FUNCTION "F_PressDemoCycleEnd" : Bool   // FC169, SCL
{ S7_Optimized_Access := 'TRUE' }
VERSION : 0.1
// stored: AutoNumber true, IsIECCheckEnabled false, SetENOAutomatically false, UDAEnableTagReadback false
   VAR_IN_OUT
      Seq : "FRK_SequenceCtx";
      Cycle : "ST_PressDemoCycle";
      Core : "FRK_Core";
      Unit : "FRK_Unit";
      Status : "ST_ModuleStatus";
      Part : "ST_PartContext";
      AlarmLog : "FRK_AlarmLog";
   END_VAR
   VAR_TEMP
      Written : Bool;
   END_VAR
BEGIN

   IF "FRK_SeqOnce"(Seq := #Seq, Enable := TRUE, Token := #Seq.Step) THEN
       #Cycle.CycleCompleted := TRUE;
       IF #Cycle.PartDispositioned THEN
           #Cycle.PartDispositioned := FALSE;
       ELSE
           #Written := "FRK_PartProcessed"(Core := #Core, Unit := #Unit, Status := #Status, Part := #Part, AlarmLog := #AlarmLog, Verdict := 1, Reason := 0);
           IF NOT #Written AND #Unit.CarrierIndex = 0 AND #Unit.Good < UDINT#4294967295 THEN
               #Unit.Good := #Unit.Good + 1;
           END_IF;
       END_IF;
       #Cycle.PartInMachine := FALSE;
       "FRK_SeqCycleEnd"(Seq := #Seq);
   END_IF;
   IF #Unit.StopReq THEN
       "FRK_Complete"(Core := #Core,
                      Status := #Status);
       "FRK_SeqComplete"(Seq := #Seq);
       #F_PressDemoCycleEnd := FALSE;
   ELSE
       #F_PressDemoCycleEnd := #Core.Exec <> 3;
   END_IF;
END_FUNCTION

FUNCTION_BLOCK "FB_LD_PressDemoHome"   // FB7, LAD
{ S7_Optimized_Access := 'TRUE' }
VERSION : 0.1
// stored: AutoNumber true, IsIECCheckEnabled false, IsRetainMemResEnabled false, MemoryReserve 100, SetENOAutomatically false, UDAEnableTagReadback false
   VAR_INPUT
      Run { ExternalWritable := 'False'} : Bool;
      Reset { ExternalWritable := 'False'} : Bool;
      OwnerIndex { ExternalWritable := 'False'} : DInt;
      Delta { ExternalWritable := 'False'} : Time;
   END_VAR
   VAR_IN_OUT
      PressRam : "FB_CylinderCM";
      Door : "FB_CylinderCM";
      PartSlide : "FB_CylinderCM";
   END_VAR
   VAR
      Seq { ExternalWritable := 'False'} : "FRK_SequenceCtx";
      Row1 { ExternalWritable := 'False'} : "FRK_SequenceRow";
      Row2 { ExternalWritable := 'False'} : "FRK_SequenceRow";
      Row3 { ExternalWritable := 'False'} : "FRK_SequenceRow";
      Row4 { ExternalWritable := 'False'} : "FRK_SequenceRow";
      At0 { ExternalAccessible := 'False'; ExternalVisible := 'False'; ExternalWritable := 'False'} : Bool;
      At900 { ExternalAccessible := 'False'; ExternalVisible := 'False'; ExternalWritable := 'False'} : Bool;
      At910 { ExternalAccessible := 'False'; ExternalVisible := 'False'; ExternalWritable := 'False'} : Bool;
      At999 { ExternalAccessible := 'False'; ExternalVisible := 'False'; ExternalWritable := 'False'} : Bool;
      Ready1 { ExternalAccessible := 'False'; ExternalVisible := 'False'; ExternalWritable := 'False'} : Bool;
      Ready2 { ExternalAccessible := 'False'; ExternalVisible := 'False'; ExternalWritable := 'False'} : Bool;
      Ready3 { ExternalAccessible := 'False'; ExternalVisible := 'False'; ExternalWritable := 'False'} : Bool;
      Ready4 { ExternalAccessible := 'False'; ExternalVisible := 'False'; ExternalWritable := 'False'} : Bool;
      Ready5 { ExternalAccessible := 'False'; ExternalVisible := 'False'; ExternalWritable := 'False'} : Bool;
      Advance { ExternalAccessible := 'False'; ExternalVisible := 'False'; ExternalWritable := 'False'} : Bool;
   END_VAR
BEGIN

REGION Network 1
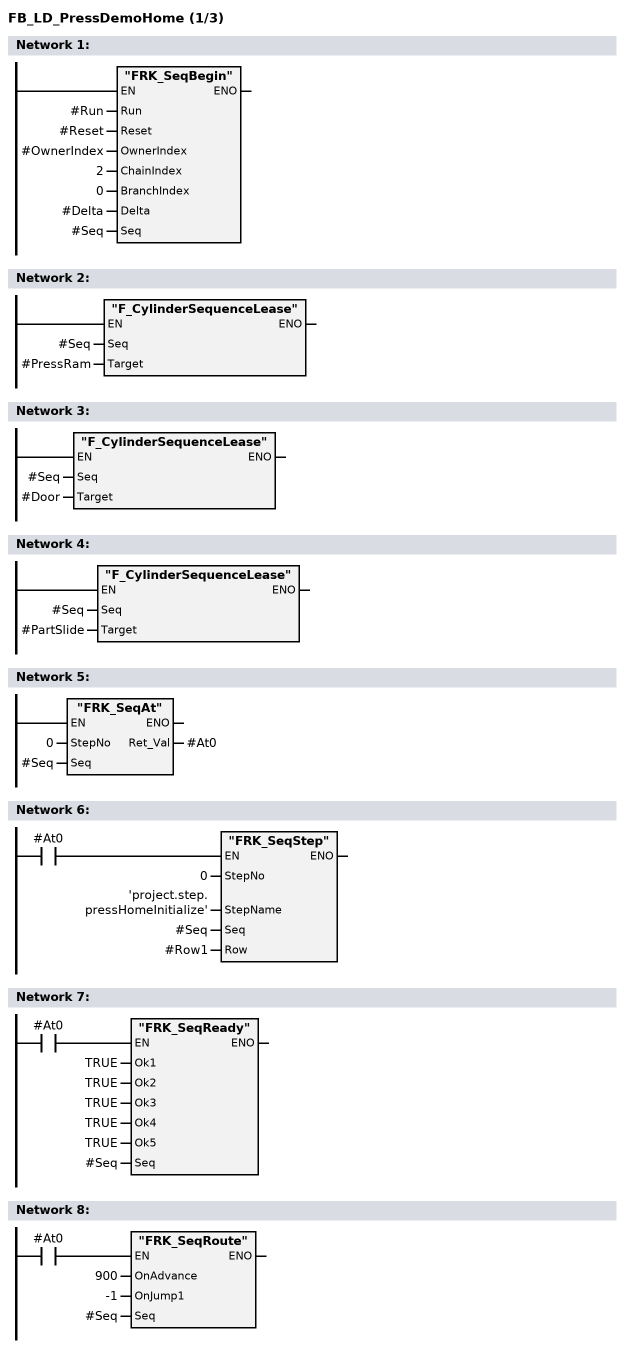
   RUNG wire#powerrail
      "FRK_SeqBegin"(Run := #Run, Reset := #Reset, OwnerIndex := #OwnerIndex, ChainIndex := 2, BranchIndex := 0, Delta := #Delta, Seq := #Seq)
   END_RUNG
   // the same network as SCL:
   "FRK_SeqBegin"(Run := #Run,
                  Reset := #Reset,
                  OwnerIndex := #OwnerIndex,
                  ChainIndex := 2,
                  BranchIndex := 0,
                  Delta := #Delta,
                  Seq := #Seq);
END_REGION

REGION Network 2
   RUNG wire#powerrail
      "F_CylinderSequenceLease"(Seq := #Seq, Target := #PressRam)
   END_RUNG
   // the same network as SCL:
   "F_CylinderSequenceLease"(Seq := #Seq, Target := #PressRam);
END_REGION

REGION Network 3
   RUNG wire#powerrail
      "F_CylinderSequenceLease"(Seq := #Seq, Target := #Door)
   END_RUNG
   // the same network as SCL:
   "F_CylinderSequenceLease"(Seq := #Seq, Target := #Door);
END_REGION

REGION Network 4
   RUNG wire#powerrail
      "F_CylinderSequenceLease"(Seq := #Seq, Target := #PartSlide)
   END_RUNG
   // the same network as SCL:
   "F_CylinderSequenceLease"(Seq := #Seq, Target := #PartSlide);
END_REGION

REGION Network 5
   RUNG wire#powerrail
      "FRK_SeqAt"(StepNo := 0, Seq := #Seq, Ret_Val => #At0)
   END_RUNG
   // the same network as SCL:
   #At0 := "FRK_SeqAt"(StepNo := 0, Seq := #Seq);
END_REGION

REGION Network 6
   RUNG wire#powerrail
      Contact( #At0 )
      "FRK_SeqStep"(StepNo := 0, StepName := 'project.step.pressHomeInitialize', Seq := #Seq, Row := #Row1)
   END_RUNG
   // the same network as SCL:
   IF #At0 THEN
       "FRK_SeqStep"(StepNo := 0, StepName := 'project.step.pressHomeInitialize', Seq := #Seq, Row := #Row1);
   END_IF;
END_REGION

REGION Network 7
   RUNG wire#powerrail
      Contact( #At0 )
      "FRK_SeqReady"(Ok1 := TRUE, Ok2 := TRUE, Ok3 := TRUE, Ok4 := TRUE, Ok5 := TRUE, Seq := #Seq)
   END_RUNG
   // the same network as SCL:
   IF #At0 THEN
       "FRK_SeqReady"(Ok1 := TRUE, Ok2 := TRUE, Ok3 := TRUE, Ok4 := TRUE, Ok5 := TRUE, Seq := #Seq);
   END_IF;
END_REGION

REGION Network 8
   RUNG wire#powerrail
      Contact( #At0 )
      "FRK_SeqRoute"(OnAdvance := 900, OnJump1 := -1, Seq := #Seq)
   END_RUNG
   // the same network as SCL:
   IF #At0 THEN "FRK_SeqRoute"(OnAdvance := 900, OnJump1 := -1, Seq := #Seq); END_IF;
END_REGION

REGION Network 9
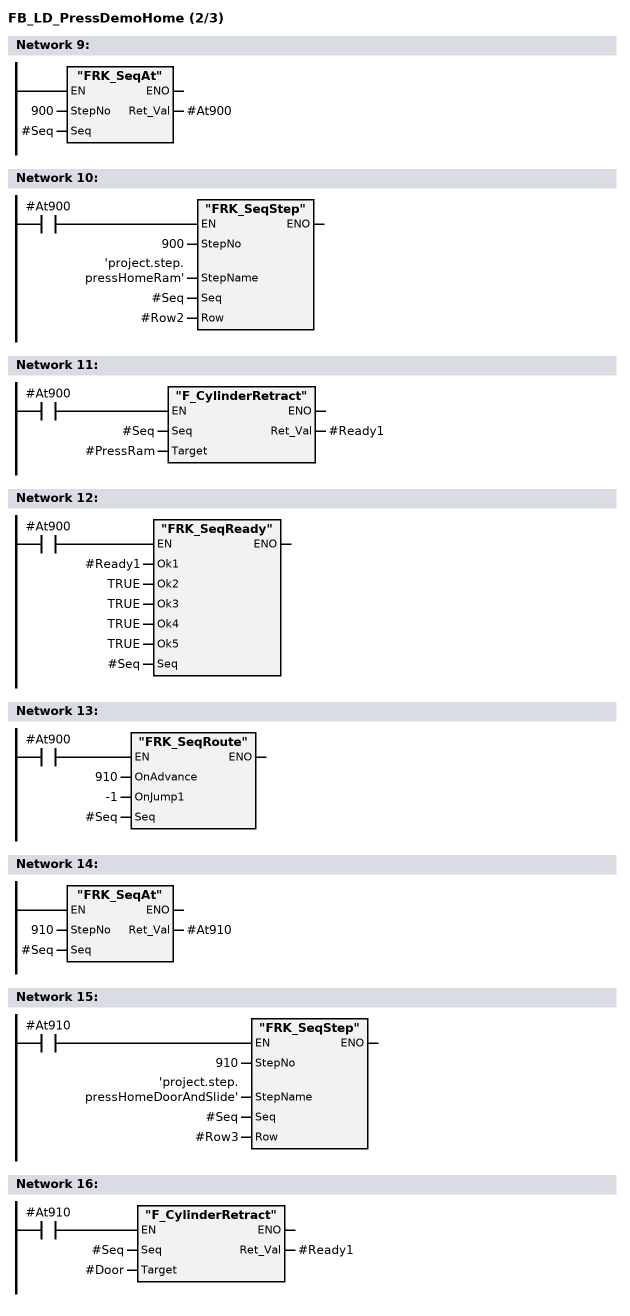
   RUNG wire#powerrail
      "FRK_SeqAt"(StepNo := 900, Seq := #Seq, Ret_Val => #At900)
   END_RUNG
   // the same network as SCL:
   #At900 := "FRK_SeqAt"(StepNo := 900, Seq := #Seq);
END_REGION

REGION Network 10
   RUNG wire#powerrail
      Contact( #At900 )
      "FRK_SeqStep"(StepNo := 900, StepName := 'project.step.pressHomeRam', Seq := #Seq, Row := #Row2)
   END_RUNG
   // the same network as SCL:
   IF #At900 THEN
       "FRK_SeqStep"(StepNo := 900, StepName := 'project.step.pressHomeRam', Seq := #Seq, Row := #Row2);
   END_IF;
END_REGION

REGION Network 11
   RUNG wire#powerrail
      Contact( #At900 )
      "F_CylinderRetract"(Seq := #Seq, Target := #PressRam, Ret_Val => #Ready1)
   END_RUNG
   // the same network as SCL:
   IF #At900 THEN #Ready1 := "F_CylinderRetract"(Seq := #Seq, Target := #PressRam); END_IF;
END_REGION

REGION Network 12
   RUNG wire#powerrail
      Contact( #At900 )
      "FRK_SeqReady"(Ok1 := #Ready1, Ok2 := TRUE, Ok3 := TRUE, Ok4 := TRUE, Ok5 := TRUE, Seq := #Seq)
   END_RUNG
   // the same network as SCL:
   IF #At900 THEN
       "FRK_SeqReady"(Ok1 := #Ready1, Ok2 := TRUE, Ok3 := TRUE, Ok4 := TRUE, Ok5 := TRUE, Seq := #Seq);
   END_IF;
END_REGION

REGION Network 13
   RUNG wire#powerrail
      Contact( #At900 )
      "FRK_SeqRoute"(OnAdvance := 910, OnJump1 := -1, Seq := #Seq)
   END_RUNG
   // the same network as SCL:
   IF #At900 THEN "FRK_SeqRoute"(OnAdvance := 910, OnJump1 := -1, Seq := #Seq); END_IF;
END_REGION

REGION Network 14
   RUNG wire#powerrail
      "FRK_SeqAt"(StepNo := 910, Seq := #Seq, Ret_Val => #At910)
   END_RUNG
   // the same network as SCL:
   #At910 := "FRK_SeqAt"(StepNo := 910, Seq := #Seq);
END_REGION

REGION Network 15
   RUNG wire#powerrail
      Contact( #At910 )
      "FRK_SeqStep"(StepNo := 910, StepName := 'project.step.pressHomeDoorAndSlide', Seq := #Seq, Row := #Row3)
   END_RUNG
   // the same network as SCL:
   IF #At910 THEN
       "FRK_SeqStep"(StepNo := 910, StepName := 'project.step.pressHomeDoorAndSlide', Seq := #Seq, Row := #Row3);
   END_IF;
END_REGION

REGION Network 16
   RUNG wire#powerrail
      Contact( #At910 )
      "F_CylinderRetract"(Seq := #Seq, Target := #Door, Ret_Val => #Ready1)
   END_RUNG
   // the same network as SCL:
   IF #At910 THEN #Ready1 := "F_CylinderRetract"(Seq := #Seq, Target := #Door); END_IF;
END_REGION

REGION Network 17
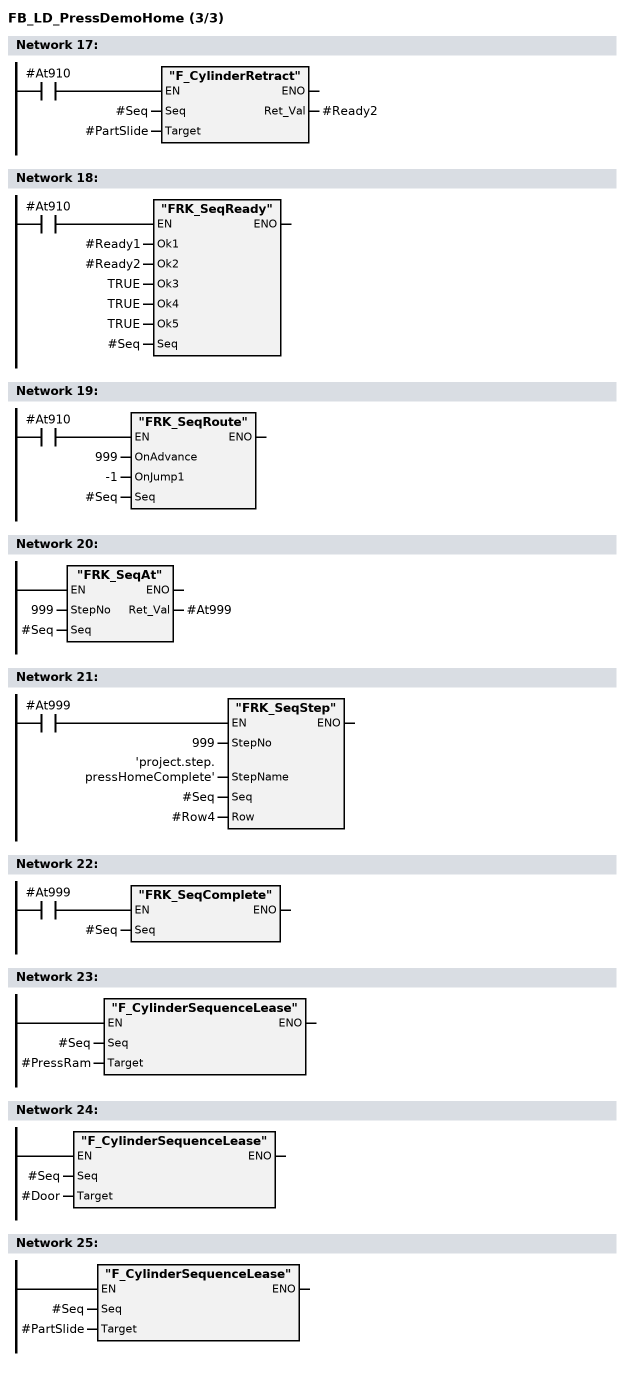
   RUNG wire#powerrail
      Contact( #At910 )
      "F_CylinderRetract"(Seq := #Seq, Target := #PartSlide, Ret_Val => #Ready2)
   END_RUNG
   // the same network as SCL:
   IF #At910 THEN #Ready2 := "F_CylinderRetract"(Seq := #Seq, Target := #PartSlide); END_IF;
END_REGION

REGION Network 18
   RUNG wire#powerrail
      Contact( #At910 )
      "FRK_SeqReady"(Ok1 := #Ready1, Ok2 := #Ready2, Ok3 := TRUE, Ok4 := TRUE, Ok5 := TRUE, Seq := #Seq)
   END_RUNG
   // the same network as SCL:
   IF #At910 THEN
       "FRK_SeqReady"(Ok1 := #Ready1, Ok2 := #Ready2, Ok3 := TRUE, Ok4 := TRUE, Ok5 := TRUE, Seq := #Seq);
   END_IF;
END_REGION

REGION Network 19
   RUNG wire#powerrail
      Contact( #At910 )
      "FRK_SeqRoute"(OnAdvance := 999, OnJump1 := -1, Seq := #Seq)
   END_RUNG
   // the same network as SCL:
   IF #At910 THEN "FRK_SeqRoute"(OnAdvance := 999, OnJump1 := -1, Seq := #Seq); END_IF;
END_REGION

REGION Network 20
   RUNG wire#powerrail
      "FRK_SeqAt"(StepNo := 999, Seq := #Seq, Ret_Val => #At999)
   END_RUNG
   // the same network as SCL:
   #At999 := "FRK_SeqAt"(StepNo := 999, Seq := #Seq);
END_REGION

REGION Network 21
   RUNG wire#powerrail
      Contact( #At999 )
      "FRK_SeqStep"(StepNo := 999, StepName := 'project.step.pressHomeComplete', Seq := #Seq, Row := #Row4)
   END_RUNG
   // the same network as SCL:
   IF #At999 THEN
       "FRK_SeqStep"(StepNo := 999, StepName := 'project.step.pressHomeComplete', Seq := #Seq, Row := #Row4);
   END_IF;
END_REGION

REGION Network 22
   RUNG wire#powerrail
      Contact( #At999 )
      "FRK_SeqComplete"(Seq := #Seq)
   END_RUNG
   // the same network as SCL:
   IF #At999 THEN "FRK_SeqComplete"(Seq := #Seq); END_IF;
END_REGION

REGION Network 23
   RUNG wire#powerrail
      "F_CylinderSequenceLease"(Seq := #Seq, Target := #PressRam)
   END_RUNG
   // the same network as SCL:
   "F_CylinderSequenceLease"(Seq := #Seq, Target := #PressRam);
END_REGION

REGION Network 24
   RUNG wire#powerrail
      "F_CylinderSequenceLease"(Seq := #Seq, Target := #Door)
   END_RUNG
   // the same network as SCL:
   "F_CylinderSequenceLease"(Seq := #Seq, Target := #Door);
END_REGION

REGION Network 25
   RUNG wire#powerrail
      "F_CylinderSequenceLease"(Seq := #Seq, Target := #PartSlide)
   END_RUNG
   // the same network as SCL:
   "F_CylinderSequenceLease"(Seq := #Seq, Target := #PartSlide);
END_REGION
END_FUNCTION_BLOCK

FUNCTION "FRK_SeqComplete" : Void   // FC127, SCL
{ S7_Optimized_Access := 'TRUE' }
VERSION : 0.1
// stored: AutoNumber true, IsIECCheckEnabled false, SetENOAutomatically false, UDAEnableTagReadback false
   VAR_IN_OUT
      Seq : "FRK_SequenceCtx";
   END_VAR
BEGIN

   #Seq.Done := TRUE;
   #Seq.Running := FALSE;
END_FUNCTION

FUNCTION_BLOCK "FB_LD_PressDemoLoadPosition"   // FB8, LAD
{ S7_Optimized_Access := 'TRUE' }
VERSION : 0.1
// stored: AutoNumber true, IsIECCheckEnabled false, IsRetainMemResEnabled false, MemoryReserve 100, SetENOAutomatically false, UDAEnableTagReadback false
   VAR_INPUT
      Run { ExternalWritable := 'False'} : Bool;
      Reset { ExternalWritable := 'False'} : Bool;
      OwnerIndex { ExternalWritable := 'False'} : DInt;
      Delta { ExternalWritable := 'False'} : Time;
   END_VAR
   VAR_IN_OUT
      PressRam : "FB_CylinderCM";
      Door : "FB_CylinderCM";
      PartSlide : "FB_CylinderCM";
   END_VAR
   VAR
      Seq { ExternalWritable := 'False'} : "FRK_SequenceCtx";
      Row1 { ExternalWritable := 'False'} : "FRK_SequenceRow";
      Row2 { ExternalWritable := 'False'} : "FRK_SequenceRow";
      Row3 { ExternalWritable := 'False'} : "FRK_SequenceRow";
      Row4 { ExternalWritable := 'False'} : "FRK_SequenceRow";
      At240 { ExternalAccessible := 'False'; ExternalVisible := 'False'; ExternalWritable := 'False'} : Bool;
      At260 { ExternalAccessible := 'False'; ExternalVisible := 'False'; ExternalWritable := 'False'} : Bool;
      At280 { ExternalAccessible := 'False'; ExternalVisible := 'False'; ExternalWritable := 'False'} : Bool;
      At300 { ExternalAccessible := 'False'; ExternalVisible := 'False'; ExternalWritable := 'False'} : Bool;
      Ready1 { ExternalAccessible := 'False'; ExternalVisible := 'False'; ExternalWritable := 'False'} : Bool;
      Ready2 { ExternalAccessible := 'False'; ExternalVisible := 'False'; ExternalWritable := 'False'} : Bool;
      Ready3 { ExternalAccessible := 'False'; ExternalVisible := 'False'; ExternalWritable := 'False'} : Bool;
      Ready4 { ExternalAccessible := 'False'; ExternalVisible := 'False'; ExternalWritable := 'False'} : Bool;
      Ready5 { ExternalAccessible := 'False'; ExternalVisible := 'False'; ExternalWritable := 'False'} : Bool;
      Advance { ExternalAccessible := 'False'; ExternalVisible := 'False'; ExternalWritable := 'False'} : Bool;
   END_VAR
BEGIN

REGION Network 1
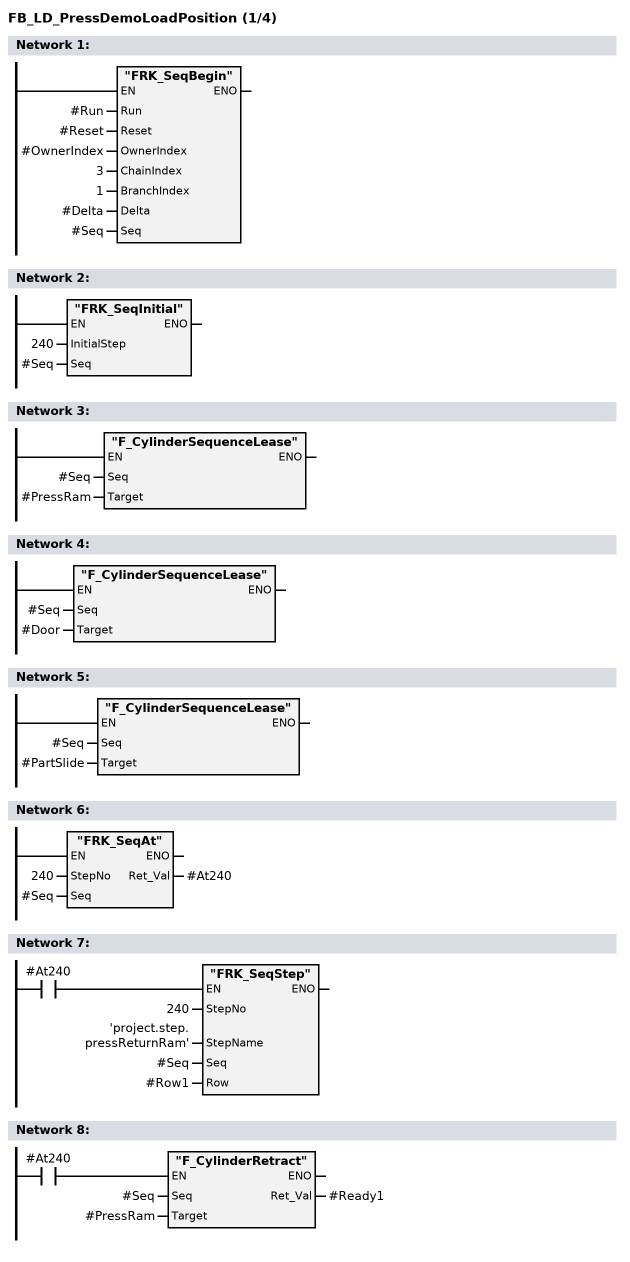
   RUNG wire#powerrail
      "FRK_SeqBegin"(Run := #Run, Reset := #Reset, OwnerIndex := #OwnerIndex, ChainIndex := 3, BranchIndex := 1, Delta := #Delta, Seq := #Seq)
   END_RUNG
   // the same network as SCL:
   "FRK_SeqBegin"(Run := #Run,
                  Reset := #Reset,
                  OwnerIndex := #OwnerIndex,
                  ChainIndex := 3,
                  BranchIndex := 1,
                  Delta := #Delta,
                  Seq := #Seq);
END_REGION

REGION Network 2
   RUNG wire#powerrail
      "FRK_SeqInitial"(InitialStep := 240, Seq := #Seq)
   END_RUNG
   // the same network as SCL:
   "FRK_SeqInitial"(InitialStep := 240, Seq := #Seq);
END_REGION

REGION Network 3
   RUNG wire#powerrail
      "F_CylinderSequenceLease"(Seq := #Seq, Target := #PressRam)
   END_RUNG
   // the same network as SCL:
   "F_CylinderSequenceLease"(Seq := #Seq, Target := #PressRam);
END_REGION

REGION Network 4
   RUNG wire#powerrail
      "F_CylinderSequenceLease"(Seq := #Seq, Target := #Door)
   END_RUNG
   // the same network as SCL:
   "F_CylinderSequenceLease"(Seq := #Seq, Target := #Door);
END_REGION

REGION Network 5
   RUNG wire#powerrail
      "F_CylinderSequenceLease"(Seq := #Seq, Target := #PartSlide)
   END_RUNG
   // the same network as SCL:
   "F_CylinderSequenceLease"(Seq := #Seq, Target := #PartSlide);
END_REGION

REGION Network 6
   RUNG wire#powerrail
      "FRK_SeqAt"(StepNo := 240, Seq := #Seq, Ret_Val => #At240)
   END_RUNG
   // the same network as SCL:
   #At240 := "FRK_SeqAt"(StepNo := 240, Seq := #Seq);
END_REGION

REGION Network 7
   RUNG wire#powerrail
      Contact( #At240 )
      "FRK_SeqStep"(StepNo := 240, StepName := 'project.step.pressReturnRam', Seq := #Seq, Row := #Row1)
   END_RUNG
   // the same network as SCL:
   IF #At240 THEN
       "FRK_SeqStep"(StepNo := 240, StepName := 'project.step.pressReturnRam', Seq := #Seq, Row := #Row1);
   END_IF;
END_REGION

REGION Network 8
   RUNG wire#powerrail
      Contact( #At240 )
      "F_CylinderRetract"(Seq := #Seq, Target := #PressRam, Ret_Val => #Ready1)
   END_RUNG
   // the same network as SCL:
   IF #At240 THEN #Ready1 := "F_CylinderRetract"(Seq := #Seq, Target := #PressRam); END_IF;
END_REGION

REGION Network 9
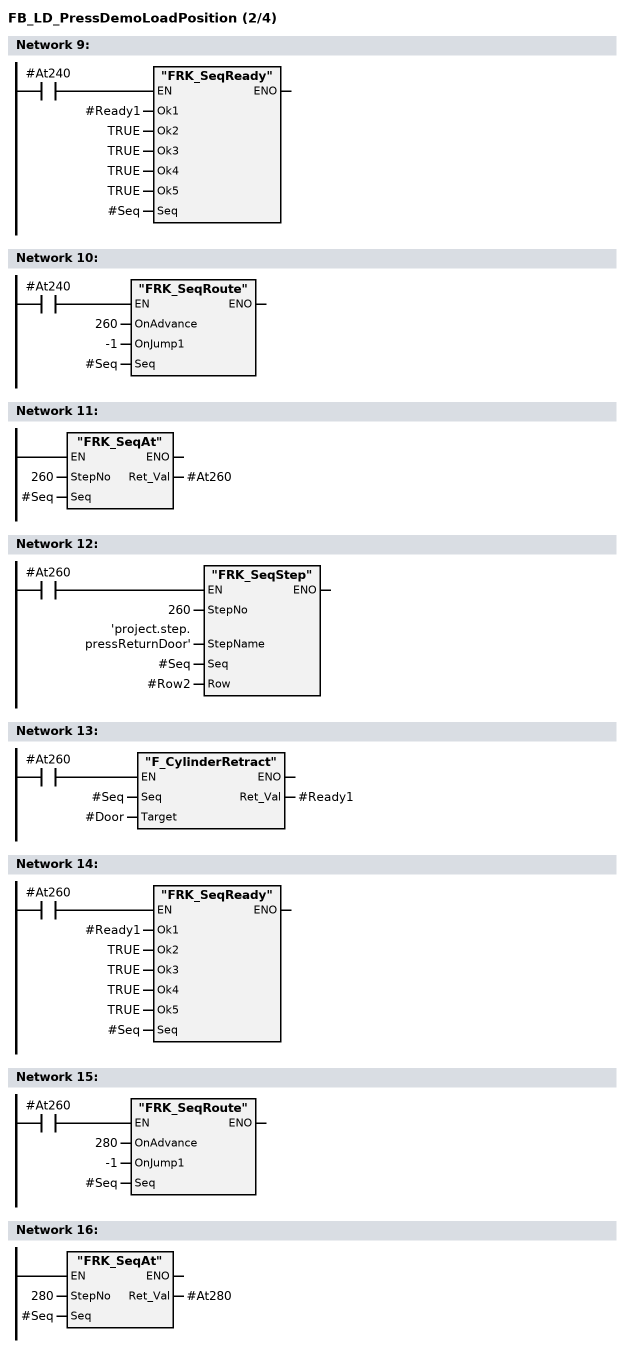
   RUNG wire#powerrail
      Contact( #At240 )
      "FRK_SeqReady"(Ok1 := #Ready1, Ok2 := TRUE, Ok3 := TRUE, Ok4 := TRUE, Ok5 := TRUE, Seq := #Seq)
   END_RUNG
   // the same network as SCL:
   IF #At240 THEN
       "FRK_SeqReady"(Ok1 := #Ready1, Ok2 := TRUE, Ok3 := TRUE, Ok4 := TRUE, Ok5 := TRUE, Seq := #Seq);
   END_IF;
END_REGION

REGION Network 10
   RUNG wire#powerrail
      Contact( #At240 )
      "FRK_SeqRoute"(OnAdvance := 260, OnJump1 := -1, Seq := #Seq)
   END_RUNG
   // the same network as SCL:
   IF #At240 THEN "FRK_SeqRoute"(OnAdvance := 260, OnJump1 := -1, Seq := #Seq); END_IF;
END_REGION

REGION Network 11
   RUNG wire#powerrail
      "FRK_SeqAt"(StepNo := 260, Seq := #Seq, Ret_Val => #At260)
   END_RUNG
   // the same network as SCL:
   #At260 := "FRK_SeqAt"(StepNo := 260, Seq := #Seq);
END_REGION

REGION Network 12
   RUNG wire#powerrail
      Contact( #At260 )
      "FRK_SeqStep"(StepNo := 260, StepName := 'project.step.pressReturnDoor', Seq := #Seq, Row := #Row2)
   END_RUNG
   // the same network as SCL:
   IF #At260 THEN
       "FRK_SeqStep"(StepNo := 260, StepName := 'project.step.pressReturnDoor', Seq := #Seq, Row := #Row2);
   END_IF;
END_REGION

REGION Network 13
   RUNG wire#powerrail
      Contact( #At260 )
      "F_CylinderRetract"(Seq := #Seq, Target := #Door, Ret_Val => #Ready1)
   END_RUNG
   // the same network as SCL:
   IF #At260 THEN #Ready1 := "F_CylinderRetract"(Seq := #Seq, Target := #Door); END_IF;
END_REGION

REGION Network 14
   RUNG wire#powerrail
      Contact( #At260 )
      "FRK_SeqReady"(Ok1 := #Ready1, Ok2 := TRUE, Ok3 := TRUE, Ok4 := TRUE, Ok5 := TRUE, Seq := #Seq)
   END_RUNG
   // the same network as SCL:
   IF #At260 THEN
       "FRK_SeqReady"(Ok1 := #Ready1, Ok2 := TRUE, Ok3 := TRUE, Ok4 := TRUE, Ok5 := TRUE, Seq := #Seq);
   END_IF;
END_REGION

REGION Network 15
   RUNG wire#powerrail
      Contact( #At260 )
      "FRK_SeqRoute"(OnAdvance := 280, OnJump1 := -1, Seq := #Seq)
   END_RUNG
   // the same network as SCL:
   IF #At260 THEN "FRK_SeqRoute"(OnAdvance := 280, OnJump1 := -1, Seq := #Seq); END_IF;
END_REGION

REGION Network 16
   RUNG wire#powerrail
      "FRK_SeqAt"(StepNo := 280, Seq := #Seq, Ret_Val => #At280)
   END_RUNG
   // the same network as SCL:
   #At280 := "FRK_SeqAt"(StepNo := 280, Seq := #Seq);
END_REGION

REGION Network 17
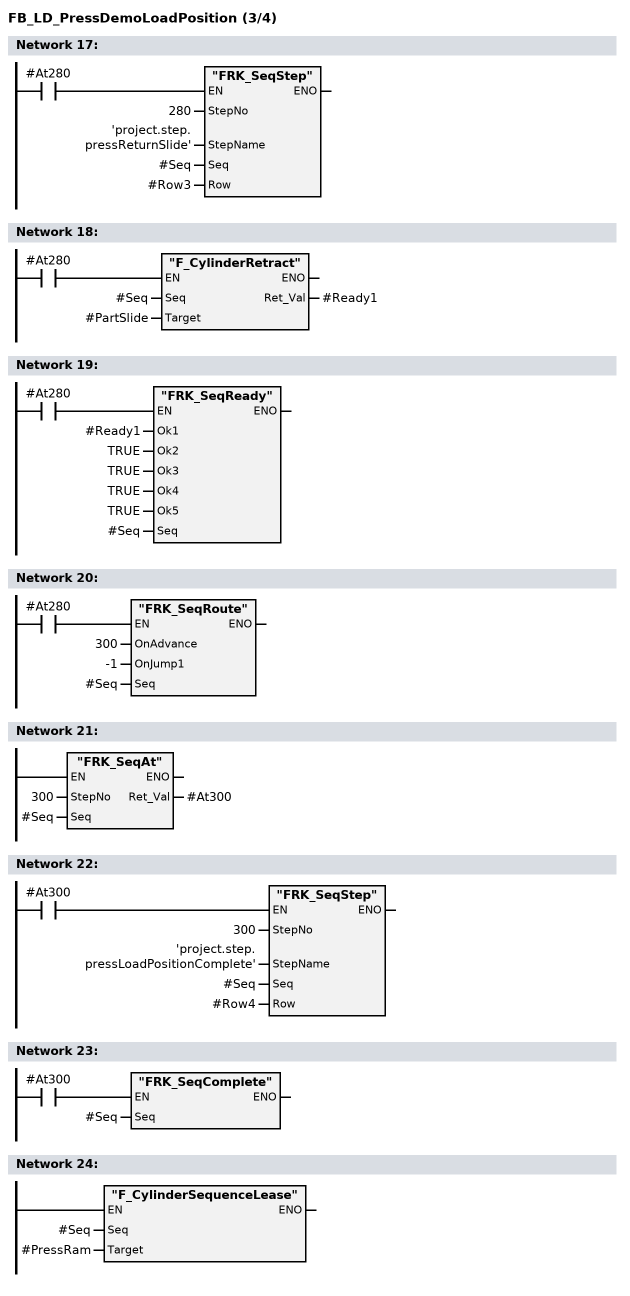
   RUNG wire#powerrail
      Contact( #At280 )
      "FRK_SeqStep"(StepNo := 280, StepName := 'project.step.pressReturnSlide', Seq := #Seq, Row := #Row3)
   END_RUNG
   // the same network as SCL:
   IF #At280 THEN
       "FRK_SeqStep"(StepNo := 280, StepName := 'project.step.pressReturnSlide', Seq := #Seq, Row := #Row3);
   END_IF;
END_REGION

REGION Network 18
   RUNG wire#powerrail
      Contact( #At280 )
      "F_CylinderRetract"(Seq := #Seq, Target := #PartSlide, Ret_Val => #Ready1)
   END_RUNG
   // the same network as SCL:
   IF #At280 THEN #Ready1 := "F_CylinderRetract"(Seq := #Seq, Target := #PartSlide); END_IF;
END_REGION

REGION Network 19
   RUNG wire#powerrail
      Contact( #At280 )
      "FRK_SeqReady"(Ok1 := #Ready1, Ok2 := TRUE, Ok3 := TRUE, Ok4 := TRUE, Ok5 := TRUE, Seq := #Seq)
   END_RUNG
   // the same network as SCL:
   IF #At280 THEN
       "FRK_SeqReady"(Ok1 := #Ready1, Ok2 := TRUE, Ok3 := TRUE, Ok4 := TRUE, Ok5 := TRUE, Seq := #Seq);
   END_IF;
END_REGION

REGION Network 20
   RUNG wire#powerrail
      Contact( #At280 )
      "FRK_SeqRoute"(OnAdvance := 300, OnJump1 := -1, Seq := #Seq)
   END_RUNG
   // the same network as SCL:
   IF #At280 THEN "FRK_SeqRoute"(OnAdvance := 300, OnJump1 := -1, Seq := #Seq); END_IF;
END_REGION

REGION Network 21
   RUNG wire#powerrail
      "FRK_SeqAt"(StepNo := 300, Seq := #Seq, Ret_Val => #At300)
   END_RUNG
   // the same network as SCL:
   #At300 := "FRK_SeqAt"(StepNo := 300, Seq := #Seq);
END_REGION

REGION Network 22
   RUNG wire#powerrail
      Contact( #At300 )
      "FRK_SeqStep"(StepNo := 300, StepName := 'project.step.pressLoadPositionComplete', Seq := #Seq, Row := #Row4)
   END_RUNG
   // the same network as SCL:
   IF #At300 THEN
       "FRK_SeqStep"(StepNo := 300, StepName := 'project.step.pressLoadPositionComplete', Seq := #Seq, Row := #Row4);
   END_IF;
END_REGION

REGION Network 23
   RUNG wire#powerrail
      Contact( #At300 )
      "FRK_SeqComplete"(Seq := #Seq)
   END_RUNG
   // the same network as SCL:
   IF #At300 THEN "FRK_SeqComplete"(Seq := #Seq); END_IF;
END_REGION

REGION Network 24
   RUNG wire#powerrail
      "F_CylinderSequenceLease"(Seq := #Seq, Target := #PressRam)
   END_RUNG
   // the same network as SCL:
   "F_CylinderSequenceLease"(Seq := #Seq, Target := #PressRam);
END_REGION

REGION Network 25
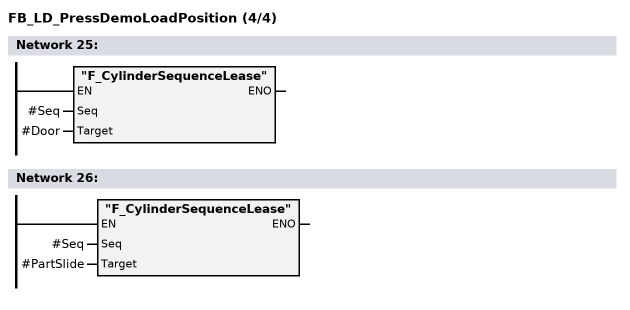
   RUNG wire#powerrail
      "F_CylinderSequenceLease"(Seq := #Seq, Target := #Door)
   END_RUNG
   // the same network as SCL:
   "F_CylinderSequenceLease"(Seq := #Seq, Target := #Door);
END_REGION

REGION Network 26
   RUNG wire#powerrail
      "F_CylinderSequenceLease"(Seq := #Seq, Target := #PartSlide)
   END_RUNG
   // the same network as SCL:
   "F_CylinderSequenceLease"(Seq := #Seq, Target := #PartSlide);
END_REGION
END_FUNCTION_BLOCK

FUNCTION "FRK_SeqInitial" : Void   // FC135, SCL
{ S7_Optimized_Access := 'TRUE' }
VERSION : 0.1
// stored: AutoNumber true, IsIECCheckEnabled false, SetENOAutomatically false, UDAEnableTagReadback false
   VAR_INPUT
      InitialStep : DInt;
   END_VAR
   VAR_IN_OUT
      Seq : "FRK_SequenceCtx";
   END_VAR
BEGIN

   IF #Seq.Restart OR NOT #Seq.Running THEN
       #Seq.Step := #InitialStep;
       #Seq.ScanStep := #InitialStep;
   END_IF;
END_FUNCTION

FUNCTION_BLOCK "FB_LD_PressDemoRelease"   // FB9, LAD
{ S7_Optimized_Access := 'TRUE' }
VERSION : 0.1
// stored: AutoNumber true, IsIECCheckEnabled false, IsRetainMemResEnabled false, MemoryReserve 100, SetENOAutomatically false, UDAEnableTagReadback false
   VAR_INPUT
      AirPressureOk { ExternalWritable := 'False'} : Bool;
      DoorClosed { ExternalWritable := 'False'} : Bool;
      DoorHealthy { ExternalWritable := 'False'} : Bool;
      RamHealthy { ExternalWritable := 'False'} : Bool;
      SlideHealthy { ExternalWritable := 'False'} : Bool;
      SlideInside { ExternalWritable := 'False'} : Bool;
      TwoHandHeld { ExternalWritable := 'False'} : Bool;
   END_VAR
   VAR
      Conditions { ExternalWritable := 'False'} : "ST_PressDemoReleaseConditions";
      ModeStart { ExternalWritable := 'False'} : "FRK_PermCtx";
      RamExtend { ExternalWritable := 'False'} : "FRK_PermCtx";
   END_VAR
BEGIN

REGION Network 1
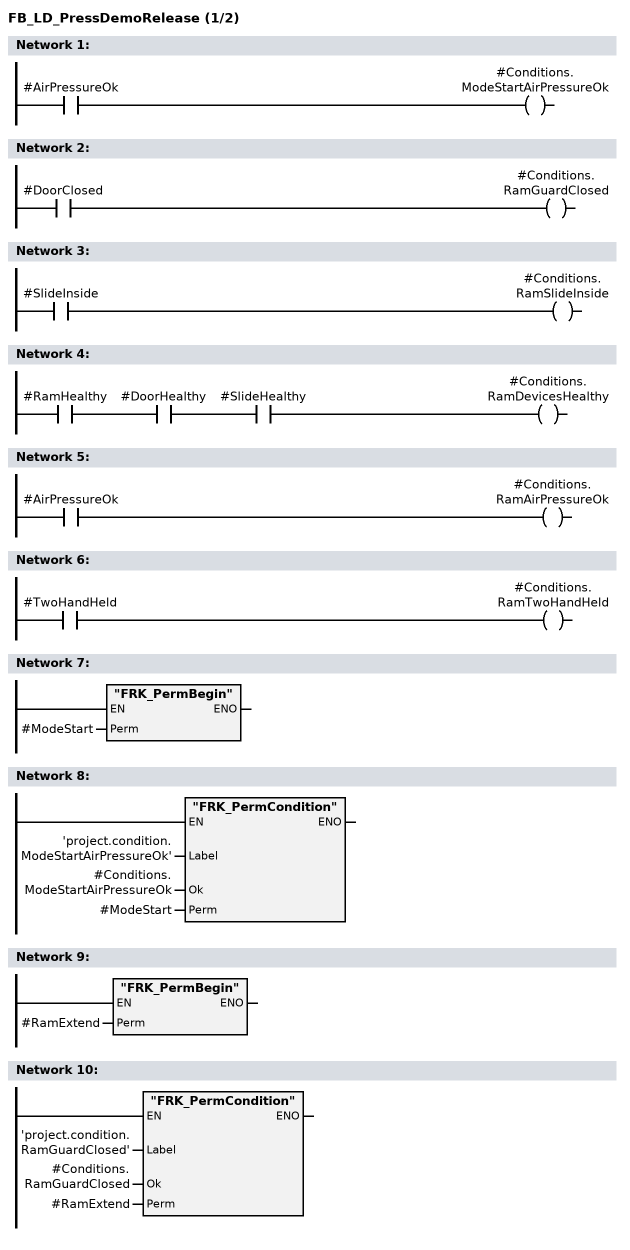
   RUNG wire#powerrail
      Contact( #AirPressureOk )
      Coil( #Conditions.ModeStartAirPressureOk )
   END_RUNG
   // the same network as SCL:
   #Conditions.ModeStartAirPressureOk := #AirPressureOk;
END_REGION

REGION Network 2
   RUNG wire#powerrail
      Contact( #DoorClosed )
      Coil( #Conditions.RamGuardClosed )
   END_RUNG
   // the same network as SCL:
   #Conditions.RamGuardClosed := #DoorClosed;
END_REGION

REGION Network 3
   RUNG wire#powerrail
      Contact( #SlideInside )
      Coil( #Conditions.RamSlideInside )
   END_RUNG
   // the same network as SCL:
   #Conditions.RamSlideInside := #SlideInside;
END_REGION

REGION Network 4
   RUNG wire#powerrail
      Contact( #RamHealthy )
      Contact( #DoorHealthy )
      Contact( #SlideHealthy )
      Coil( #Conditions.RamDevicesHealthy )
   END_RUNG
   // the same network as SCL:
   #Conditions.RamDevicesHealthy := #RamHealthy AND #DoorHealthy AND #SlideHealthy;
END_REGION

REGION Network 5
   RUNG wire#powerrail
      Contact( #AirPressureOk )
      Coil( #Conditions.RamAirPressureOk )
   END_RUNG
   // the same network as SCL:
   #Conditions.RamAirPressureOk := #AirPressureOk;
END_REGION

REGION Network 6
   RUNG wire#powerrail
      Contact( #TwoHandHeld )
      Coil( #Conditions.RamTwoHandHeld )
   END_RUNG
   // the same network as SCL:
   #Conditions.RamTwoHandHeld := #TwoHandHeld;
END_REGION

REGION Network 7
   RUNG wire#powerrail
      "FRK_PermBegin"(Perm := #ModeStart)
   END_RUNG
   // the same network as SCL:
   "FRK_PermBegin"(Perm := #ModeStart);
END_REGION

REGION Network 8
   RUNG wire#powerrail
      "FRK_PermCondition"(Label := 'project.condition.ModeStartAirPressureOk', Ok := #Conditions.ModeStartAirPressureOk, Perm := #ModeStart)
   END_RUNG
   // the same network as SCL:
   "FRK_PermCondition"(Label := 'project.condition.ModeStartAirPressureOk',
                       Ok := #Conditions.ModeStartAirPressureOk,
                       Perm := #ModeStart);
END_REGION

REGION Network 9
   RUNG wire#powerrail
      "FRK_PermBegin"(Perm := #RamExtend)
   END_RUNG
   // the same network as SCL:
   "FRK_PermBegin"(Perm := #RamExtend);
END_REGION

REGION Network 10
   RUNG wire#powerrail
      "FRK_PermCondition"(Label := 'project.condition.RamGuardClosed', Ok := #Conditions.RamGuardClosed, Perm := #RamExtend)
   END_RUNG
   // the same network as SCL:
   "FRK_PermCondition"(Label := 'project.condition.RamGuardClosed',
                       Ok := #Conditions.RamGuardClosed,
                       Perm := #RamExtend);
END_REGION

REGION Network 11
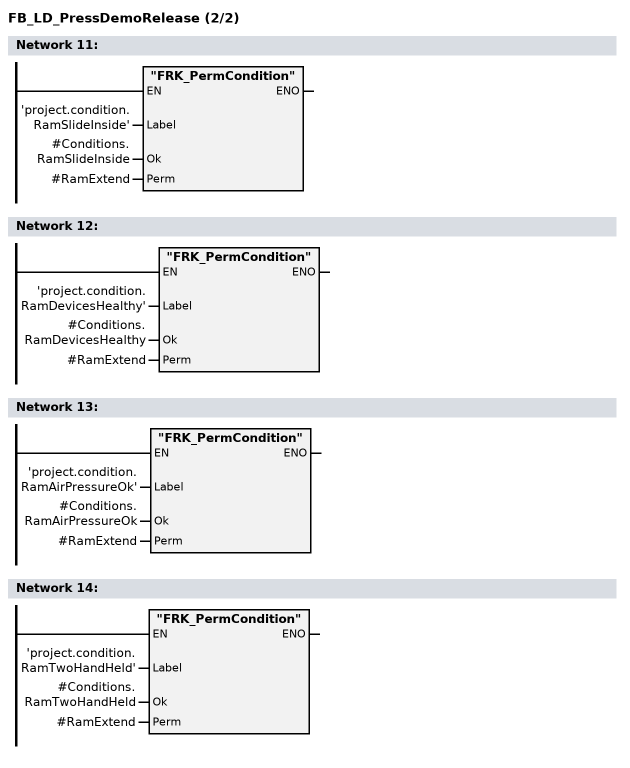
   RUNG wire#powerrail
      "FRK_PermCondition"(Label := 'project.condition.RamSlideInside', Ok := #Conditions.RamSlideInside, Perm := #RamExtend)
   END_RUNG
   // the same network as SCL:
   "FRK_PermCondition"(Label := 'project.condition.RamSlideInside',
                       Ok := #Conditions.RamSlideInside,
                       Perm := #RamExtend);
END_REGION

REGION Network 12
   RUNG wire#powerrail
      "FRK_PermCondition"(Label := 'project.condition.RamDevicesHealthy', Ok := #Conditions.RamDevicesHealthy, Perm := #RamExtend)
   END_RUNG
   // the same network as SCL:
   "FRK_PermCondition"(Label := 'project.condition.RamDevicesHealthy',
                       Ok := #Conditions.RamDevicesHealthy,
                       Perm := #RamExtend);
END_REGION

REGION Network 13
   RUNG wire#powerrail
      "FRK_PermCondition"(Label := 'project.condition.RamAirPressureOk', Ok := #Conditions.RamAirPressureOk, Perm := #RamExtend)
   END_RUNG
   // the same network as SCL:
   "FRK_PermCondition"(Label := 'project.condition.RamAirPressureOk',
                       Ok := #Conditions.RamAirPressureOk,
                       Perm := #RamExtend);
END_REGION

REGION Network 14
   RUNG wire#powerrail
      "FRK_PermCondition"(Label := 'project.condition.RamTwoHandHeld', Ok := #Conditions.RamTwoHandHeld, Perm := #RamExtend)
   END_RUNG
   // the same network as SCL:
   "FRK_PermCondition"(Label := 'project.condition.RamTwoHandHeld',
                       Ok := #Conditions.RamTwoHandHeld,
                       Perm := #RamExtend);
END_REGION
END_FUNCTION_BLOCK

FUNCTION "FRK_PermBegin" : Void   // FC122, SCL
{ S7_Optimized_Access := 'TRUE' }
VERSION : 0.1
// One collection sweep and first FALSE condition, shared by ST and LAD.
// stored: AutoNumber true, IsIECCheckEnabled false, SetENOAutomatically false, UDAEnableTagReadback false
   VAR_IN_OUT
      Perm : "FRK_PermCtx";
   END_VAR
BEGIN

   #Perm.Permit := TRUE;
   #Perm.Blocker := '';
   #Perm.Count := 0;
END_FUNCTION

FUNCTION "FRK_PermCondition" : Void   // FC123, SCL
{ S7_Optimized_Access := 'TRUE' }
VERSION : 0.1
// stored: AutoNumber true, IsIECCheckEnabled false, SetENOAutomatically false, UDAEnableTagReadback false
   VAR_INPUT
      Label : String;
      Ok : Bool;
   END_VAR
   VAR_IN_OUT
      Perm : "FRK_PermCtx";
   END_VAR
BEGIN

   #Perm.Count := #Perm.Count + 1;
   IF NOT #Ok THEN
       IF #Perm.Permit THEN
           #Perm.Blocker := #Label;
       END_IF;
       #Perm.Permit := FALSE;
   END_IF;
END_FUNCTION

FUNCTION_BLOCK "FB_PressDemoAuto"   // FB3, SCL
{ S7_Optimized_Access := 'TRUE' }
VERSION : 0.1
// stored: AutoNumber true, IsIECCheckEnabled false, IsRetainMemResEnabled false, MemoryReserve 100, SetENOAutomatically false, UDAEnableTagReadback false
   VAR_INPUT
      Run : Bool;
      Reset : Bool;
      OwnerIndex : DInt;
      Delta : Time;
      TransferSettleTime : Time;
      PartQuality : Bool;
      RequireTwoHandStart : Bool;
      SourcePath : String[80];
      PartPresent : Bool;
      AirPressureOk : Bool;
      TwoHandHeld : Bool;
      StartPulse : Bool;
      PressSettleTime : Time;
   END_VAR
   VAR_IN_OUT
      PressRam : "FB_CylinderCM";
      Door : "FB_CylinderCM";
      PartSlide : "FB_CylinderCM";
      Core : "FRK_Core";
      Unit : "FRK_Unit";
      Status : "ST_ModuleStatus";
      Part : "ST_PartContext";
      AlarmLog : "FRK_AlarmLog";
   END_VAR
   VAR
      Seq { ExternalWritable := 'False'; S7_SetPoint := 'True'} : "FRK_SequenceCtx";
      Row1 { ExternalWritable := 'False'; S7_SetPoint := 'True'} : "FRK_SequenceRow";
      Row2 { ExternalWritable := 'False'; S7_SetPoint := 'True'} : "FRK_SequenceRow";
      Row3 { ExternalWritable := 'False'; S7_SetPoint := 'True'} : "FRK_SequenceRow";
      Row4 { ExternalWritable := 'False'; S7_SetPoint := 'True'} : "FRK_SequenceRow";
      Row5 { ExternalWritable := 'False'; S7_SetPoint := 'True'} : "FRK_SequenceRow";
      Row6 { ExternalWritable := 'False'; S7_SetPoint := 'True'} : "FRK_SequenceRow";
      Row7 { ExternalWritable := 'False'; S7_SetPoint := 'True'} : "FRK_SequenceRow";
      Row8 { ExternalWritable := 'False'; S7_SetPoint := 'True'} : "FRK_SequenceRow";
      Row9 { ExternalWritable := 'False'; S7_SetPoint := 'True'} : "FRK_SequenceRow";
      Row10 { ExternalWritable := 'False'; S7_SetPoint := 'True'} : "FRK_SequenceRow";
      Row11 { ExternalWritable := 'False'; S7_SetPoint := 'True'} : "FRK_SequenceRow";
      Row12 { ExternalWritable := 'False'; S7_SetPoint := 'True'} : "FRK_SequenceRow";
      Row13 { ExternalWritable := 'False'; S7_SetPoint := 'True'} : "FRK_SequenceRow";
      Row14 { ExternalWritable := 'False'; S7_SetPoint := 'True'} : "FRK_SequenceRow";
      Row15 { ExternalWritable := 'False'; S7_SetPoint := 'True'} : "FRK_SequenceRow";
      Row16 { ExternalWritable := 'False'; S7_SetPoint := 'True'} : "FRK_SequenceRow";
      At0 { ExternalAccessible := 'False'; ExternalVisible := 'False'; ExternalWritable := 'False'} : Bool;
      At100 { ExternalAccessible := 'False'; ExternalVisible := 'False'; ExternalWritable := 'False'} : Bool;
      At110 { ExternalAccessible := 'False'; ExternalVisible := 'False'; ExternalWritable := 'False'} : Bool;
      At130 { ExternalAccessible := 'False'; ExternalVisible := 'False'; ExternalWritable := 'False'} : Bool;
      At150 { ExternalAccessible := 'False'; ExternalVisible := 'False'; ExternalWritable := 'False'} : Bool;
      At170 { ExternalAccessible := 'False'; ExternalVisible := 'False'; ExternalWritable := 'False'} : Bool;
      At180 { ExternalAccessible := 'False'; ExternalVisible := 'False'; ExternalWritable := 'False'} : Bool;
      At185 { ExternalAccessible := 'False'; ExternalVisible := 'False'; ExternalWritable := 'False'} : Bool;
      At190 { ExternalAccessible := 'False'; ExternalVisible := 'False'; ExternalWritable := 'False'} : Bool;
      At200 { ExternalAccessible := 'False'; ExternalVisible := 'False'; ExternalWritable := 'False'} : Bool;
      At210 { ExternalAccessible := 'False'; ExternalVisible := 'False'; ExternalWritable := 'False'} : Bool;
      At215 { ExternalAccessible := 'False'; ExternalVisible := 'False'; ExternalWritable := 'False'} : Bool;
      At220 { ExternalAccessible := 'False'; ExternalVisible := 'False'; ExternalWritable := 'False'} : Bool;
      At230 { ExternalAccessible := 'False'; ExternalVisible := 'False'; ExternalWritable := 'False'} : Bool;
      At240 { ExternalAccessible := 'False'; ExternalVisible := 'False'; ExternalWritable := 'False'} : Bool;
      At999 { ExternalAccessible := 'False'; ExternalVisible := 'False'; ExternalWritable := 'False'} : Bool;
      Ready1 { ExternalAccessible := 'False'; ExternalVisible := 'False'; ExternalWritable := 'False'} : Bool;
      Ready2 { ExternalAccessible := 'False'; ExternalVisible := 'False'; ExternalWritable := 'False'} : Bool;
      Ready3 { ExternalAccessible := 'False'; ExternalVisible := 'False'; ExternalWritable := 'False'} : Bool;
      Ready4 { ExternalAccessible := 'False'; ExternalVisible := 'False'; ExternalWritable := 'False'} : Bool;
      Ready5 { ExternalAccessible := 'False'; ExternalVisible := 'False'; ExternalWritable := 'False'} : Bool;
      Advance { ExternalAccessible := 'False'; ExternalVisible := 'False'; ExternalWritable := 'False'} : Bool;
      Cycle { ExternalAccessible := 'False'; ExternalVisible := 'False'; ExternalWritable := 'False'; S7_SetPoint := 'True'} : "ST_PressDemoCycle";
      LoadPosition { ExternalAccessible := 'False'; ExternalVisible := 'False'; ExternalWritable := 'False'; S7_SetPoint := 'True'} : "FB_PressDemoLoadPosition";
      LoadDone { ExternalAccessible := 'False'; ExternalVisible := 'False'; ExternalWritable := 'False'} : Bool;
      LoadActive { ExternalAccessible := 'False'; ExternalVisible := 'False'; ExternalWritable := 'False'} : Bool;
   END_VAR
BEGIN

   "FRK_SeqBegin"(Run := #Run,
                  Reset := #Reset,
                  OwnerIndex := #OwnerIndex,
                  ChainIndex := 1,
                  BranchIndex := 0,
                  Delta := #Delta,
                  Seq := #Seq);
   "FRK_SeqStart"(Seq := #Seq,
                  StartPulse := #StartPulse);
   "F_PressDemoReset"(Seq := #Seq,
                      Cycle := #Cycle);
   #LoadActive := "FRK_SeqSubActive"(Seq := #Seq, Run := #Run, StepNo := 240);
   #LoadDone := "F_PressDemoLoadPosition"(Target := #LoadPosition, Run := #LoadActive, Reset := #Seq.Restart, OwnerIndex := #OwnerIndex, Delta := #Delta, PressRam := #PressRam, Door := #Door, PartSlide := #PartSlide);
   "F_CylinderSequenceLease"(Seq := #Seq,
                             Target := #PressRam);
   "F_CylinderSequenceLease"(Seq := #Seq,
                             Target := #Door);
   "F_CylinderSequenceLease"(Seq := #Seq,
                             Target := #PartSlide);
   "FRK_SeqOwnerStatus"(Seq := #Seq,
                        Core := #Core,
                        Status := #Status);
   "FRK_SeqSubStatus"(Seq := #Seq,
                      Child := #LoadPosition.Seq);
   CASE #Seq.ScanStep OF
       0:
           IF #Seq.Running AND NOT #Seq.Error THEN
               "FRK_SeqStep"(StepNo := 0,
                             StepName := 'project.step.pressAutoInitialize',
                             Seq := #Seq,
                             Row := #Row1);
               "FRK_SeqReady"(Seq := #Seq,
                              Ok1 := TRUE,
                              Ok2 := TRUE,
                              Ok3 := TRUE,
                              Ok4 := TRUE,
                              Ok5 := TRUE);
               "FRK_SeqRoute"(Seq := #Seq,
                              OnAdvance := 100,
                              OnJump1 := -1);
           END_IF;
       100:
           IF #Seq.Running AND NOT #Seq.Error THEN
               "FRK_SeqStep"(StepNo := 100,
                             StepName := 'project.step.pressAwaitTwoHand',
                             Seq := #Seq,
                             Row := #Row2);
               #Ready5 := "F_PressDemoAwaitCycle"(Seq := #Seq, Cycle := #Cycle, Core := #Core, Unit := #Unit, Status := #Status, Part := #Part, AlarmLog := #AlarmLog, PartPresent := #PartPresent, PartQuality := #PartQuality, AirPressureOk := #AirPressureOk, RequireTwoHandStart := #RequireTwoHandStart);
               "FRK_SeqReady"(Seq := #Seq,
                              Ok1 := #Ready5,
                              Ok2 := TRUE,
                              Ok3 := TRUE,
                              Ok4 := TRUE,
                              Ok5 := TRUE);
               "FRK_SeqRoute"(Seq := #Seq,
                              OnAdvance := 110,
                              OnJump1 := -1);
           END_IF;
       110:
           IF #Seq.Running AND NOT #Seq.Error THEN
               "FRK_SeqStep"(StepNo := 110,
                             StepName := 'project.step.pressRamUp',
                             Seq := #Seq,
                             Row := #Row3);
               #Ready1 := "F_CylinderRetract"(Seq := #Seq, Target := #PressRam);
               "FRK_SeqReady"(Seq := #Seq,
                              Ok1 := #Ready1,
                              Ok2 := TRUE,
                              Ok3 := TRUE,
                              Ok4 := TRUE,
                              Ok5 := TRUE);
               "FRK_SeqRoute"(Seq := #Seq,
                              OnAdvance := 130,
                              OnJump1 := -1);
           END_IF;
       130:
           IF #Seq.Running AND NOT #Seq.Error THEN
               "FRK_SeqStep"(StepNo := 130,
                             StepName := 'project.step.pressDoorOpen',
                             Seq := #Seq,
                             Row := #Row4);
               #Ready1 := "F_CylinderRetract"(Seq := #Seq, Target := #Door);
               "FRK_SeqReady"(Seq := #Seq,
                              Ok1 := #Ready1,
                              Ok2 := TRUE,
                              Ok3 := TRUE,
                              Ok4 := TRUE,
                              Ok5 := TRUE);
               "FRK_SeqRoute"(Seq := #Seq,
                              OnAdvance := 150,
                              OnJump1 := -1);
           END_IF;
       150:
           IF #Seq.Running AND NOT #Seq.Error THEN
               "FRK_SeqStep"(StepNo := 150,
                             StepName := 'project.step.pressSlideInside',
                             Seq := #Seq,
                             Row := #Row5);
               #Ready1 := "F_CylinderExtend"(Seq := #Seq, Target := #PartSlide);
               "F_PressDemoStarted"(Seq := #Seq,
                                    Unit := #Unit,
                                    Status := #Status,
                                    Part := #Part,
                                    AlarmLog := #AlarmLog);
               "FRK_SeqReady"(Seq := #Seq,
                              Ok1 := #Ready1,
                              Ok2 := TRUE,
                              Ok3 := TRUE,
                              Ok4 := TRUE,
                              Ok5 := TRUE);
               "FRK_SeqRoute"(Seq := #Seq,
                              OnAdvance := 170,
                              OnJump1 := -1);
           END_IF;
       170:
           IF #Seq.Running AND NOT #Seq.Error THEN
               "FRK_SeqStep"(StepNo := 170,
                             StepName := 'project.step.pressTransferSettle',
                             Seq := #Seq,
                             Row := #Row6);
               #Ready1 := "FRK_SeqDelay"(Seq := #Seq, PT := #TransferSettleTime, Delta := #Delta, Permit := TRUE);
               "FRK_SeqReady"(Seq := #Seq,
                              Ok1 := #Ready1,
                              Ok2 := TRUE,
                              Ok3 := TRUE,
                              Ok4 := TRUE,
                              Ok5 := TRUE);
               "FRK_SeqRoute"(Seq := #Seq,
                              OnAdvance := 180,
                              OnJump1 := -1);
           END_IF;
       180:
           IF #Seq.Running AND NOT #Seq.Error THEN
               "FRK_SeqStep"(StepNo := 180,
                             StepName := 'project.step.pressDoorClose',
                             Seq := #Seq,
                             Row := #Row7);
               #Ready1 := "F_CylinderExtend"(Seq := #Seq, Target := #Door);
               "F_PressDemoDoorClose"(Seq := #Seq,
                                      Closed := #Ready1,
                                      TwoHandHeld := #TwoHandHeld,
                                      RequireTwoHandStart := #RequireTwoHandStart,
                                      SourcePath := #SourcePath,
                                      AlarmLog := #AlarmLog);
               "FRK_SeqRoute"(Seq := #Seq,
                              OnAdvance := 200,
                              OnJump1 := 185);
           END_IF;
       185:
           IF #Seq.Running AND NOT #Seq.Error THEN
               "FRK_SeqStep"(StepNo := 185,
                             StepName := 'project.step.pressDoorReopen',
                             Seq := #Seq,
                             Row := #Row8);
               #Ready1 := "F_CylinderRetract"(Seq := #Seq, Target := #Door);
               "FRK_SeqReady"(Seq := #Seq,
                              Ok1 := #Ready1,
                              Ok2 := TRUE,
                              Ok3 := TRUE,
                              Ok4 := TRUE,
                              Ok5 := TRUE);
               "FRK_SeqRoute"(Seq := #Seq,
                              OnAdvance := 190,
                              OnJump1 := -1);
           END_IF;
       190:
           IF #Seq.Running AND NOT #Seq.Error THEN
               "FRK_SeqStep"(StepNo := 190,
                             StepName := 'project.step.pressSlideOutsideAfterAbort',
                             Seq := #Seq,
                             Row := #Row9);
               #Ready1 := "F_CylinderRetract"(Seq := #Seq, Target := #PartSlide);
               "F_PressDemoClearStart"(Seq := #Seq,
                                       Complete := #Ready1);
               "FRK_SeqReady"(Seq := #Seq,
                              Ok1 := #Ready1,
                              Ok2 := TRUE,
                              Ok3 := TRUE,
                              Ok4 := TRUE,
                              Ok5 := TRUE);
               "FRK_SeqRoute"(Seq := #Seq,
                              OnAdvance := 100,
                              OnJump1 := -1);
           END_IF;
       200:
           IF #Seq.Running AND NOT #Seq.Error THEN
               "FRK_SeqStep"(StepNo := 200,
                             StepName := 'project.step.pressRamDown',
                             Seq := #Seq,
                             Row := #Row10);
               #Ready1 := "F_CylinderExtendHandled"(Seq := #Seq, Target := #PressRam);
               "F_PressDemoRamResult"(Seq := #Seq,
                                      Reached := #Ready1,
                                      Cycle := #Cycle,
                                      AlarmLog := #AlarmLog);
               "FRK_SeqRoute"(Seq := #Seq,
                              OnAdvance := 220,
                              OnJump1 := 210);
           END_IF;
       210:
           IF #Seq.Running AND NOT #Seq.Error THEN
               "FRK_SeqStep"(StepNo := 210,
                             StepName := 'project.step.pressNotReachedConfirm',
                             Seq := #Seq,
                             Row := #Row11);
               #Ready5 := "F_PressDemoConfirmScrap"(Seq := #Seq, SourcePath := #SourcePath, AlarmLog := #AlarmLog);
               "FRK_SeqReady"(Seq := #Seq,
                              Ok1 := #Ready5,
                              Ok2 := TRUE,
                              Ok3 := TRUE,
                              Ok4 := TRUE,
                              Ok5 := TRUE);
               "FRK_SeqRoute"(Seq := #Seq,
                              OnAdvance := 215,
                              OnJump1 := -1);
           END_IF;
       215:
           IF #Seq.Running AND NOT #Seq.Error THEN
               "FRK_SeqStep"(StepNo := 215,
                             StepName := 'project.step.pressScrapPart',
                             Seq := #Seq,
                             Row := #Row12);
               #Ready5 := "F_PressDemoScrap"(Seq := #Seq, Cycle := #Cycle, Core := #Core, Unit := #Unit, Status := #Status, Part := #Part, AlarmLog := #AlarmLog);
               "FRK_SeqReady"(Seq := #Seq,
                              Ok1 := #Ready5,
                              Ok2 := TRUE,
                              Ok3 := TRUE,
                              Ok4 := TRUE,
                              Ok5 := TRUE);
               "FRK_SeqRoute"(Seq := #Seq,
                              OnAdvance := 240,
                              OnJump1 := -1);
           END_IF;
       220:
           IF #Seq.Running AND NOT #Seq.Error THEN
               "FRK_SeqStep"(StepNo := 220,
                             StepName := 'project.step.pressDwell',
                             Seq := #Seq,
                             Row := #Row13);
               #Ready5 := "F_PressDemoDwell"(Seq := #Seq, TwoHandHeld := #TwoHandHeld, RequireTwoHandStart := #RequireTwoHandStart, PT := #PressSettleTime, Delta := #Delta, PressRam := #PressRam);
               "FRK_SeqReady"(Seq := #Seq,
                              Ok1 := #Ready5,
                              Ok2 := TRUE,
                              Ok3 := TRUE,
                              Ok4 := TRUE,
                              Ok5 := TRUE);
               "FRK_SeqRoute"(Seq := #Seq,
                              OnAdvance := 230,
                              OnJump1 := -1);
           END_IF;
       230:
           IF #Seq.Running AND NOT #Seq.Error THEN
               "FRK_SeqStep"(StepNo := 230,
                             StepName := 'project.step.pressRecordResult',
                             Seq := #Seq,
                             Row := #Row14);
               #Ready5 := "F_PressDemoRecord"(Seq := #Seq, Dwell := #PressSettleTime, Core := #Core, Status := #Status, Part := #Part);
               "FRK_SeqReady"(Seq := #Seq,
                              Ok1 := #Ready5,
                              Ok2 := TRUE,
                              Ok3 := TRUE,
                              Ok4 := TRUE,
                              Ok5 := TRUE);
               "FRK_SeqRoute"(Seq := #Seq,
                              OnAdvance := 240,
                              OnJump1 := -1);
           END_IF;
       240:
           IF #Seq.Running AND NOT #Seq.Error THEN
               "FRK_SeqStep"(StepNo := 240,
                             StepName := 'project.step.pressReturnToLoad',
                             Seq := #Seq,
                             Row := #Row15);
               #Ready1 := "FRK_SeqAwait"(Seq := #Seq, Label := 'project.condition.LoadDone', Ok := #LoadDone);
               "FRK_SeqReady"(Seq := #Seq,
                              Ok1 := #Ready1,
                              Ok2 := TRUE,
                              Ok3 := TRUE,
                              Ok4 := TRUE,
                              Ok5 := TRUE);
               "FRK_SeqRoute"(Seq := #Seq,
                              OnAdvance := 999,
                              OnJump1 := -1);
           END_IF;
       999:
           IF #Seq.Running AND NOT #Seq.Error THEN
               "FRK_SeqStep"(StepNo := 999,
                             StepName := 'project.step.pressAutoComplete',
                             Seq := #Seq,
                             Row := #Row16);
               #Ready5 := "F_PressDemoCycleEnd"(Seq := #Seq, Cycle := #Cycle, Core := #Core, Unit := #Unit, Status := #Status, Part := #Part, AlarmLog := #AlarmLog);
               "FRK_SeqReady"(Seq := #Seq,
                              Ok1 := #Ready5,
                              Ok2 := TRUE,
                              Ok3 := TRUE,
                              Ok4 := TRUE,
                              Ok5 := TRUE);
               "FRK_SeqRoute"(Seq := #Seq,
                              OnAdvance := 100,
                              OnJump1 := -1);
           END_IF;
       ELSE
           #Seq.Error := TRUE;
           #Seq.ErrorDiagnostic.ReasonCode := 10001;
           #Seq.ErrorDiagnostic.Description := WSTRING#'project.sequence.invalidStep';
   END_CASE;
   "F_CylinderSequenceLease"(Seq := #Seq,
                             Target := #PressRam);
   "F_CylinderSequenceLease"(Seq := #Seq,
                             Target := #Door);
   "F_CylinderSequenceLease"(Seq := #Seq,
                             Target := #PartSlide);
   "FRK_SeqOwnerStatus"(Seq := #Seq,
                        Core := #Core,
                        Status := #Status);
   "FRK_SeqSubStatus"(Seq := #Seq,
                      Child := #LoadPosition.Seq);
END_FUNCTION_BLOCK

FUNCTION_BLOCK "FB_PressDemoHardwareDriver"   // FB14, SCL
{ S7_Optimized_Access := 'TRUE' }
VERSION : 0.1
// stored: AutoNumber true, IsIECCheckEnabled false, IsRetainMemResEnabled false, MemoryReserve 100, SetENOAutomatically false, UDAEnableTagReadback false
   VAR_INPUT
      ReadInputs { ExternalAccessible := 'False'; ExternalVisible := 'False'; ExternalWritable := 'False'} : Bool;
   END_VAR
BEGIN

   IF #ReadInputs THEN
       "GDB_FraktalHal".Data.PressDemo.Process.PartPresent := "GDB_PressDemoIO".PartPresent;
       "GDB_FraktalHal".Data.PressDemo.Process.PartQuality := "GDB_PressDemoIO".PartQuality;
       "GDB_FraktalHal".Data.PressDemo.Process.AirPressureOk := "GDB_PressDemoIO".AirPressureOk;
       "GDB_FraktalHal".Data.PressDemo.Process.TwoHandHeld := "GDB_PressDemoIO".TwoHandHeld;
       "GDB_FraktalHal".Data.PressDemo.Process.StartPulse := "GDB_PressDemoIO".StartPulse;
       "GDB_FraktalHal".Data.PressDemo.PressRam.FeedbackExtended := "GDB_PressDemoIO".RamExtended;
       "GDB_FraktalHal".Data.PressDemo.PressRam.FeedbackRetracted := "GDB_PressDemoIO".RamRetracted;
       "GDB_FraktalHal".Data.PressDemo.Door.FeedbackExtended := "GDB_PressDemoIO".DoorClosed;
       "GDB_FraktalHal".Data.PressDemo.Door.FeedbackRetracted := "GDB_PressDemoIO".DoorOpen;
       "GDB_FraktalHal".Data.PressDemo.PartSlide.FeedbackExtended := "GDB_PressDemoIO".SlideInside;
       "GDB_FraktalHal".Data.PressDemo.PartSlide.FeedbackRetracted := "GDB_PressDemoIO".SlideOutside;
   ELSE
       "GDB_PressDemoIO".RamExtend := "GDB_FraktalHal".Data.PressDemo.PressRam.CoilExtend;
       "GDB_PressDemoIO".RamRetract := "GDB_FraktalHal".Data.PressDemo.PressRam.CoilRetract;
       "GDB_PressDemoIO".DoorClose := "GDB_FraktalHal".Data.PressDemo.Door.CoilExtend;
       "GDB_PressDemoIO".DoorRelease := "GDB_FraktalHal".Data.PressDemo.Door.CoilRetract;
       "GDB_PressDemoIO".SlideExtend := "GDB_FraktalHal".Data.PressDemo.PartSlide.CoilExtend;
       "GDB_PressDemoIO".SlideRetract := "GDB_FraktalHal".Data.PressDemo.PartSlide.CoilRetract;
   END_IF;
END_FUNCTION_BLOCK

FUNCTION_BLOCK "FB_PressDemoHome"   // FB4, SCL
{ S7_Optimized_Access := 'TRUE' }
VERSION : 0.1
// stored: AutoNumber true, IsIECCheckEnabled false, IsRetainMemResEnabled false, MemoryReserve 100, SetENOAutomatically false, UDAEnableTagReadback false
   VAR_INPUT
      Run : Bool;
      Reset : Bool;
      OwnerIndex : DInt;
      Delta : Time;
   END_VAR
   VAR_IN_OUT
      PressRam : "FB_CylinderCM";
      Door : "FB_CylinderCM";
      PartSlide : "FB_CylinderCM";
   END_VAR
   VAR
      Seq { ExternalWritable := 'False'; S7_SetPoint := 'True'} : "FRK_SequenceCtx";
      Row1 { ExternalWritable := 'False'; S7_SetPoint := 'True'} : "FRK_SequenceRow";
      Row2 { ExternalWritable := 'False'; S7_SetPoint := 'True'} : "FRK_SequenceRow";
      Row3 { ExternalWritable := 'False'; S7_SetPoint := 'True'} : "FRK_SequenceRow";
      Row4 { ExternalWritable := 'False'; S7_SetPoint := 'True'} : "FRK_SequenceRow";
      At0 { ExternalAccessible := 'False'; ExternalVisible := 'False'; ExternalWritable := 'False'} : Bool;
      At900 { ExternalAccessible := 'False'; ExternalVisible := 'False'; ExternalWritable := 'False'} : Bool;
      At910 { ExternalAccessible := 'False'; ExternalVisible := 'False'; ExternalWritable := 'False'} : Bool;
      At999 { ExternalAccessible := 'False'; ExternalVisible := 'False'; ExternalWritable := 'False'} : Bool;
      Ready1 { ExternalAccessible := 'False'; ExternalVisible := 'False'; ExternalWritable := 'False'} : Bool;
      Ready2 { ExternalAccessible := 'False'; ExternalVisible := 'False'; ExternalWritable := 'False'} : Bool;
      Ready3 { ExternalAccessible := 'False'; ExternalVisible := 'False'; ExternalWritable := 'False'} : Bool;
      Ready4 { ExternalAccessible := 'False'; ExternalVisible := 'False'; ExternalWritable := 'False'} : Bool;
      Ready5 { ExternalAccessible := 'False'; ExternalVisible := 'False'; ExternalWritable := 'False'} : Bool;
      Advance { ExternalAccessible := 'False'; ExternalVisible := 'False'; ExternalWritable := 'False'} : Bool;
   END_VAR
BEGIN

   "FRK_SeqBegin"(Run := #Run,
                  Reset := #Reset,
                  OwnerIndex := #OwnerIndex,
                  ChainIndex := 2,
                  BranchIndex := 0,
                  Delta := #Delta,
                  Seq := #Seq);
   "F_CylinderSequenceLease"(Seq := #Seq,
                             Target := #PressRam);
   "F_CylinderSequenceLease"(Seq := #Seq,
                             Target := #Door);
   "F_CylinderSequenceLease"(Seq := #Seq,
                             Target := #PartSlide);
   CASE #Seq.ScanStep OF
       0:
           IF #Seq.Running AND NOT #Seq.Error THEN
               "FRK_SeqStep"(StepNo := 0,
                             StepName := 'project.step.pressHomeInitialize',
                             Seq := #Seq,
                             Row := #Row1);
               "FRK_SeqReady"(Seq := #Seq,
                              Ok1 := TRUE,
                              Ok2 := TRUE,
                              Ok3 := TRUE,
                              Ok4 := TRUE,
                              Ok5 := TRUE);
               "FRK_SeqRoute"(Seq := #Seq,
                              OnAdvance := 900,
                              OnJump1 := -1);
           END_IF;
       900:
           IF #Seq.Running AND NOT #Seq.Error THEN
               "FRK_SeqStep"(StepNo := 900,
                             StepName := 'project.step.pressHomeRam',
                             Seq := #Seq,
                             Row := #Row2);
               #Ready1 := "F_CylinderRetract"(Seq := #Seq, Target := #PressRam);
               "FRK_SeqReady"(Seq := #Seq,
                              Ok1 := #Ready1,
                              Ok2 := TRUE,
                              Ok3 := TRUE,
                              Ok4 := TRUE,
                              Ok5 := TRUE);
               "FRK_SeqRoute"(Seq := #Seq,
                              OnAdvance := 910,
                              OnJump1 := -1);
           END_IF;
       910:
           IF #Seq.Running AND NOT #Seq.Error THEN
               "FRK_SeqStep"(StepNo := 910,
                             StepName := 'project.step.pressHomeDoorAndSlide',
                             Seq := #Seq,
                             Row := #Row3);
               #Ready1 := "F_CylinderRetract"(Seq := #Seq, Target := #Door);
               #Ready2 := "F_CylinderRetract"(Seq := #Seq, Target := #PartSlide);
               "FRK_SeqReady"(Seq := #Seq,
                              Ok1 := #Ready1,
                              Ok2 := #Ready2,
                              Ok3 := TRUE,
                              Ok4 := TRUE,
                              Ok5 := TRUE);
               "FRK_SeqRoute"(Seq := #Seq,
                              OnAdvance := 999,
                              OnJump1 := -1);
           END_IF;
       999:
           IF #Seq.Running AND NOT #Seq.Error THEN
               "FRK_SeqStep"(StepNo := 999,
                             StepName := 'project.step.pressHomeComplete',
                             Seq := #Seq,
                             Row := #Row4);
               "FRK_SeqComplete"(Seq := #Seq);
           END_IF;
       ELSE
           #Seq.Error := TRUE;
           #Seq.ErrorDiagnostic.ReasonCode := 10001;
           #Seq.ErrorDiagnostic.Description := WSTRING#'project.sequence.invalidStep';
   END_CASE;
   "F_CylinderSequenceLease"(Seq := #Seq,
                             Target := #PressRam);
   "F_CylinderSequenceLease"(Seq := #Seq,
                             Target := #Door);
   "F_CylinderSequenceLease"(Seq := #Seq,
                             Target := #PartSlide);
END_FUNCTION_BLOCK

FUNCTION "FRK_AccessAudit" : Void   // FC45, SCL
{ S7_Optimized_Access := 'TRUE' }
VERSION : 0.1
// stored: AutoNumber true, IsIECCheckEnabled false, SetENOAutomatically false, UDAEnableTagReadback false
   VAR_INPUT
      What : WString;
      Who : String;
      SourcePath : WString;
   END_VAR
   VAR_IN_OUT
      AlarmLog : "FRK_AlarmLog";
   END_VAR
   VAR_TEMP
      Description : WString[480];
   END_VAR
BEGIN

   #Description := CONCAT(IN1 := #What, IN2 := WSTRING#': ');
   #Description := CONCAT(IN1 := #Description, IN2 := STRING_TO_WSTRING(#Who));
   "FRK_AlarmMessage"(AlarmLog := #AlarmLog,
                      Reason := 0,
                      Description := #Description,
                      SourcePath := #SourcePath);
END_FUNCTION

FUNCTION "FRK_AccessCancel" : Void   // FC40, SCL
{ S7_Optimized_Access := 'TRUE' }
VERSION : 0.1
// stored: AutoNumber true, IsIECCheckEnabled false, SetENOAutomatically false, UDAEnableTagReadback false
   VAR_IN_OUT
      Access : "FRK_Access";
   END_VAR
   VAR_TEMP
      Index : DInt;
   END_VAR
BEGIN

   #Access.LoginBusy := FALSE;
   #Access.CandidateUser := '';
   #Access.CandidateLevel := 0;
   #Access.Round := 0;
   FOR #Index := 0 TO 15 DO
       #Access.Salt[#Index] := 0;
   END_FOR;
   FOR #Index := 0 TO 31 DO
       #Access.Digest[#Index] := 0;
       #Access.Expected[#Index] := 0;
   END_FOR;
END_FUNCTION

FUNCTION "FRK_AccessCrcByte" : DWord   // FC48, SCL
{ S7_Optimized_Access := 'TRUE' }
VERSION : 0.1
// Reference-1500 LOCAL_RETAIN adapter. No sessions or plaintext credentials.
//  CRC-32 arithmetic comes from Core F_Crc32; encoding is binding-local, versioned.
// stored: AutoNumber true, IsIECCheckEnabled false, SetENOAutomatically false, UDAEnableTagReadback false
   VAR_INPUT
      Previous : DWord;
      Value : Byte;
   END_VAR
   VAR_TEMP
      BitIndex : Int;
      Work : DWord;
   END_VAR
BEGIN

   #Work := #Previous XOR BYTE_TO_DWORD(#Value);
   FOR #BitIndex := 0 TO 7 DO
       IF (#Work AND DWORD#1) <> 0 THEN
           #Work := SHR(IN := #Work, N := 1) XOR DWORD#16#EDB88320;
       ELSE
           #Work := SHR(IN := #Work, N := 1);
       END_IF;
   END_FOR;
   #FRK_AccessCrcByte := #Work;
END_FUNCTION

FUNCTION "FRK_AccessCrcNumber" : DWord   // FC49, SCL
{ S7_Optimized_Access := 'TRUE' }
VERSION : 0.1
// stored: AutoNumber true, IsIECCheckEnabled false, SetENOAutomatically false, UDAEnableTagReadback false
   VAR_INPUT
      Previous : DWord;
      Value : UDInt;
   END_VAR
   VAR_TEMP
      Index : Int;
      Work : DWord;
   END_VAR
BEGIN

   #Work := #Previous;
   FOR #Index := 0 TO 3 DO
       #Work := "FRK_AccessCrcByte"(Previous := #Work, Value := DWORD_TO_BYTE(SHR(IN := UDINT_TO_DWORD(#Value), N := INT_TO_UINT(#Index * 8))));
   END_FOR;
   #FRK_AccessCrcNumber := #Work;
END_FUNCTION

FUNCTION "FRK_AccessCyclic" : Void   // FC46, SCL
{ S7_Optimized_Access := 'TRUE' }
VERSION : 0.1
// stored: AutoNumber true, IsIECCheckEnabled false, SetENOAutomatically false, UDAEnableTagReadback false
   VAR_INPUT
      Startup : Bool;
      SourcePath : WString;
   END_VAR
   VAR_IN_OUT
      Access : "FRK_Access";
      AlarmLog : "FRK_AlarmLog";
      Revision : UDInt;
   END_VAR
   VAR_TEMP
      Data : Array[0..47] of Byte;
      Index : DInt;
      Difference : Byte;
      HashOk : Bool;
   END_VAR
BEGIN

   #Access.LoginTimeoutMs := 6000;
   IF #Startup THEN
       "FRK_AccessLogout"(Access := #Access);
       #Access.LoginResultSequence := 0;
   END_IF;
   IF #Access.ProviderGeneration <> "FRK_LocalUsers".Generation OR NOT "FRK_AccessStorage".UsersReady THEN
       IF #Access.CurrentLevel > 0 THEN
           "FRK_AccessAudit"(AlarmLog := #AlarmLog,
                             What := WSTRING#'std.audit.autoLogout',
                             Who := #Access.CurrentUser,
                             SourcePath := #SourcePath);
           "FRK_AccessDropSession"(Access := #Access);
           #Revision := "FRK_ConfigRevision"(Previous := #Revision);
       END_IF;
       IF #Access.LoginBusy THEN
           #Access.CandidateLevel := 0;
       END_IF;
       #Access.ProviderGeneration := "FRK_LocalUsers".Generation;
   END_IF;
   IF #Access.CurrentLevel > 0 AND #Access.Policy.SessionTimeout > T#0ms THEN
       IF "FRK_Elapsed"(NewMs := "FRK_Clock".NowMs, OldMs := #Access.LastActivity) >= DINT_TO_UDINT(TIME_TO_DINT(#Access.Policy.SessionTimeout)) THEN
           "FRK_AccessAudit"(AlarmLog := #AlarmLog,
                             What := WSTRING#'std.audit.autoLogout',
                             Who := #Access.CurrentUser,
                             SourcePath := #SourcePath);
           // Expiring the old session does not discard a separately committed
           // credential attempt. Explicit logout cancels both.
           "FRK_AccessDropSession"(Access := #Access);
           #Revision := "FRK_ConfigRevision"(Previous := #Revision);
       END_IF;
   END_IF;
   IF NOT #Access.LoginBusy THEN
       RETURN;
   END_IF;
   // One compression per active scan; never run all PIN rounds in one scan.
   FOR #Index := 0 TO 31 DO
       #Data[#Index] := #Access.Digest[#Index];
   END_FOR;
   FOR #Index := 0 TO 15 DO
       #Data[32 + #Index] := #Access.Salt[#Index];
   END_FOR;
   #HashOk := "FRK_Sha256Pin"(Data := #Data, Size := 48, Digest := #Access.Digest);
   FOR #Index := 0 TO 47 DO
       #Data[#Index] := 0;
   END_FOR;
   #Access.Round := #Access.Round + 1;
   IF NOT #HashOk OR "FRK_Elapsed"(NewMs := "FRK_Clock".NowMs, OldMs := #Access.LoginSince) >= #Access.LoginTimeoutMs THEN
       #Access.CandidateLevel := 0;
   ELSIF #Access.Round < 256 THEN
       RETURN;
   END_IF;
   #Difference := 0;
   FOR #Index := 0 TO 31 DO
       #Difference := #Difference OR (#Access.Digest[#Index] XOR #Access.Expected[#Index]);
   END_FOR;
   #Access.LoginFailed := #Difference <> 0 OR #Access.CandidateLevel = 0 OR NOT #Access.ProviderEnabled OR NOT "FRK_AccessStorage".UsersReady OR #Access.CandidateGeneration <> "FRK_LocalUsers".Generation;
   IF #Access.LoginFailed THEN
       "FRK_AccessAudit"(AlarmLog := #AlarmLog,
                         What := WSTRING#'std.audit.loginFailed',
                         Who := #Access.CandidateUser,
                         SourcePath := #SourcePath);
   ELSE
       #Access.CurrentUser := #Access.CandidateUser;
       #Access.CurrentLevel := #Access.CandidateLevel;
       #Access.LastActivity := "FRK_Clock".NowMs;
       #Access.SessionGeneration := "FRK_AccessNext"(Previous := #Access.SessionGeneration);
       #Revision := "FRK_ConfigRevision"(Previous := #Revision);
       "FRK_AccessAudit"(AlarmLog := #AlarmLog,
                         What := WSTRING#'std.audit.login',
                         Who := #Access.CurrentUser,
                         SourcePath := #SourcePath);
   END_IF;
   #Access.LoginResultSequence := #Access.LoginSequence;
   "FRK_AccessCancel"(Access := #Access);
END_FUNCTION

FUNCTION "FRK_AccessDropSession" : Void   // FC42, SCL
{ S7_Optimized_Access := 'TRUE' }
VERSION : 0.1
// stored: AutoNumber true, IsIECCheckEnabled false, SetENOAutomatically false, UDAEnableTagReadback false
   VAR_IN_OUT
      Access : "FRK_Access";
   END_VAR
BEGIN

   #Access.CurrentLevel := 0;
   #Access.CurrentUser := '';
   #Access.LoginFailed := FALSE;
   #Access.SessionGeneration := "FRK_AccessNext"(Previous := #Access.SessionGeneration);
END_FUNCTION

FUNCTION "FRK_AccessFinish" : Void   // FC47, SCL
{ S7_Optimized_Access := 'TRUE' }
VERSION : 0.1
// stored: AutoNumber true, IsIECCheckEnabled false, SetENOAutomatically false, UDAEnableTagReadback false
   VAR_INPUT
      Unit : "FRK_Unit";
      Response : "ST_HmiResponse";
      SourcePath : WString;
   END_VAR
   VAR_IN_OUT
      Access : "FRK_Access";
      AlarmLog : "FRK_AlarmLog";
      Revision : UDInt;
   END_VAR
   VAR_TEMP
      What : WString[160];
      AuditPath : WString[255];
   END_VAR
BEGIN

   IF NOT #Unit.RequestPending THEN
       RETURN;
   END_IF;
   CASE #Unit.Request.Kind OF
       23, 15,
       16, 17,
       1:
           RETURN;
       2:
           "FRK_AccessAudit"(AlarmLog := #AlarmLog,
                             What := WSTRING#'std.audit.logout',
                             Who := #Unit.RequestUser,
                             SourcePath := #SourcePath);
           #Revision := "FRK_ConfigRevision"(Previous := #Revision);
           RETURN;
       ELSE
           #What := WSTRING#'std.audit.accessDenied';
   END_CASE;
   IF #Response.Accepted THEN
       #What := WSTRING#'std.audit.operatorAction';
       IF #Access.CurrentLevel > 0 THEN
           #Access.LastActivity := "FRK_Clock".NowMs;
       END_IF;
       IF #Unit.Request.Kind = 24 OR #Unit.Request.Kind = 25 THEN
           #Revision := "FRK_ConfigRevision"(Previous := #Revision);
       END_IF;
   END_IF;
   #AuditPath := #SourcePath;
   IF #Unit.Request.Kind = 11 THEN
       IF #Response.Accepted THEN
           #AuditPath := #Unit.Request.TargetPath;
       END_IF;
       IF #Response.Accepted THEN
           #What := WSTRING#'std.audit.manualCommandAccepted';
       ELSE
           #What := WSTRING#'std.audit.manualCommandRejected';
       END_IF;
   END_IF;
   #What := CONCAT(IN1 := #What, IN2 := WSTRING#' kind=');
   #What := CONCAT(IN1 := #What, IN2 := DINT_TO_WSTRING(#Unit.Request.Kind));
   #What := CONCAT(IN1 := #What, IN2 := WSTRING#' value=');
   #What := CONCAT(IN1 := #What, IN2 := DINT_TO_WSTRING(#Unit.Request.IntValue));
   "FRK_AccessAudit"(AlarmLog := #AlarmLog,
                     What := #What,
                     Who := #Unit.RequestUser,
                     SourcePath := #AuditPath);
END_FUNCTION

FUNCTION "FRK_AccessLogin" : Void   // FC44, SCL
{ S7_Optimized_Access := 'TRUE' }
VERSION : 0.1
// stored: AutoNumber true, IsIECCheckEnabled false, SetENOAutomatically false, UDAEnableTagReadback false
   VAR_INPUT
      User : String;
      Secret : String;
      Sequence : UDInt;
   END_VAR
   VAR_IN_OUT
      Access : "FRK_Access";
   END_VAR
   VAR_TEMP
      Data : Array[0..47] of Byte;
      Index : DInt;
      Slot : DInt;
      Size : Int;
      HashOk : Bool;
   END_VAR
BEGIN

   "FRK_AccessCancel"(Access := #Access);
   #Access.LoginFailed := FALSE;
   #Access.LoginSequence := #Sequence;
   #Access.CandidateGeneration := "FRK_LocalUsers".Generation;
   #Access.LoginSince := "FRK_Clock".NowMs;
   #Access.LoginTimeoutMs := 6000;
   #Access.CandidateUser := #User;
   // Unknown users execute the same bounded work with a dummy salt/digest.
   IF #Access.ProviderEnabled AND "FRK_AccessStorage".UsersReady AND "FRK_LocalUsers".Count >= 0 AND "FRK_LocalUsers".Count <= 16 THEN
       FOR #Slot := 1 TO "FRK_LocalUsers".Count DO
           IF #User <> '' AND "FRK_LocalUsers".Rows[#Slot].User = #User THEN
               IF "FRK_LocalUsers".Rows[#Slot].Level >= 1 AND "FRK_LocalUsers".Rows[#Slot].Level <= 4 THEN
                   #Access.CandidateLevel := "FRK_LocalUsers".Rows[#Slot].Level;
                   #Access.Salt := "FRK_LocalUsers".Rows[#Slot].Salt;
                   #Access.Expected := "FRK_LocalUsers".Rows[#Slot].PinHash;
               END_IF;
               EXIT;
           END_IF;
       END_FOR;
   END_IF;
   FOR #Index := 0 TO 47 DO
       #Data[#Index] := 0;
   END_FOR;
   FOR #Index := 0 TO 15 DO
       #Data[#Index] := #Access.Salt[#Index];
   END_FOR;
   #Size := LEN(#Secret);
   IF #Size > 32 THEN
       #Size := 0;
       #Access.CandidateLevel := 0;
   END_IF;
   FOR #Index := 1 TO #Size DO
       #Data[15 + #Index] := CHAR_TO_BYTE(#Secret[#Index]);
   END_FOR;
   #HashOk := "FRK_Sha256Pin"(Data := #Data, Size := 16 + INT_TO_DINT(#Size), Digest := #Access.Digest);
   FOR #Index := 0 TO 47 DO
       #Data[#Index] := 0;
   END_FOR;
   #Access.LoginBusy := #HashOk;
END_FUNCTION

FUNCTION "FRK_AccessLogout" : Void   // FC41, SCL
{ S7_Optimized_Access := 'TRUE' }
VERSION : 0.1
// stored: AutoNumber true, IsIECCheckEnabled false, SetENOAutomatically false, UDAEnableTagReadback false
   VAR_IN_OUT
      Access : "FRK_Access";
   END_VAR
BEGIN

   "FRK_AccessCancel"(Access := #Access);
   "FRK_AccessDropSession"(Access := #Access);
END_FUNCTION

FUNCTION "FRK_AccessNext" : UDInt   // FC43, SCL
{ S7_Optimized_Access := 'TRUE' }
VERSION : 0.1
// stored: AutoNumber true, IsIECCheckEnabled false, SetENOAutomatically false, UDAEnableTagReadback false
   VAR_INPUT
      Previous : UDInt;
   END_VAR
BEGIN

   IF #Previous = UDINT#4294967295 THEN
       #FRK_AccessNext := 1;
   ELSE
       #FRK_AccessNext := #Previous + 1;
   END_IF;
END_FUNCTION

FUNCTION "FRK_AccessPersist" : Void   // FC60, SCL
{ S7_Optimized_Access := 'TRUE' }
VERSION : 0.1
// stored: AutoNumber true, IsIECCheckEnabled false, SetENOAutomatically false, UDAEnableTagReadback false
   VAR_INPUT
      Unit : "FRK_Unit";
      SourcePath : WString;
   END_VAR
   VAR_IN_OUT
      Access : "FRK_Access";
      Response : "ST_HmiResponse";
      AlarmLog : "FRK_AlarmLog";
   END_VAR
   VAR_TEMP
      Diag : "ST_Diagnostic";
      Accepted : Bool;
   END_VAR
BEGIN

   IF #Unit.RequestPending AND #Unit.Request.Kind = 31 AND #Access.PolicyLost THEN
       // Explicit ENGINEER acknowledgement accepts the restrictive fallback.
       #Response.Accepted := #Access.CurrentLevel >= 3 AND #Access.PolicySlot > 0;
       IF #Response.Accepted THEN
           "FRK_AccessPolicySave"(Access := #Access,
                                  Scope := WSTRING_TO_STRING(#SourcePath));
           #Access.PolicyLost := FALSE;
           #Response.Diagnostic := WSTRING#'';
       ELSE
           #Response.Diagnostic := WSTRING#'std.error.configRestoreAckRefused';
       END_IF;
   ELSIF #Unit.RequestPending AND #Response.Accepted AND NOT #Access.PolicyLost AND (#Unit.Request.Kind = 24 OR #Unit.Request.Kind = 25) THEN
       "FRK_AccessPolicySave"(Access := #Access,
                              Scope := WSTRING_TO_STRING(#SourcePath));
   END_IF;
   IF #Access.PolicyLost AND #Access.PolicyLossAlarm = 0 THEN
       #Diag := "FRK_UnitScratch".EmptyDiagnostic;
       #Diag.ReasonCode := 2040;
       #Diag.Description := WSTRING#'std.error.configRestoreLost';
       #Diag.SourcePath := #SourcePath;
       #Access.PolicyLossAlarm := "FRK_AlarmRaise"(AlarmLog := #AlarmLog, Diag := #Diag, ResetClass := 0);
   ELSIF NOT #Access.PolicyLost AND #Access.PolicyLossAlarm > 0 THEN
       #Accepted := "FRK_AlarmGone"(AlarmLog := #AlarmLog, Slot := #Access.PolicyLossAlarm);
       #Access.PolicyLossAlarm := 0;
   END_IF;
   IF "FRK_AccessStorage".UsersLost AND #Access.PolicySlot > 0 AND #Access.UserLossAlarm = 0 THEN
       #Diag := "FRK_UnitScratch".EmptyDiagnostic;
       #Diag.ReasonCode := 2040;
       #Diag.Description := WSTRING#'std.error.accessRestoreLost';
       #Diag.SourcePath := #SourcePath;
       #Access.UserLossAlarm := "FRK_AlarmRaise"(AlarmLog := #AlarmLog, Diag := #Diag, ResetClass := 0);
   ELSIF NOT "FRK_AccessStorage".UsersLost AND #Access.UserLossAlarm > 0 THEN
       #Accepted := "FRK_AlarmGone"(AlarmLog := #AlarmLog, Slot := #Access.UserLossAlarm);
       #Access.UserLossAlarm := 0;
   END_IF;
END_FUNCTION

FUNCTION "FRK_AccessPolicyBoot" : Void   // FC59, SCL
{ S7_Optimized_Access := 'TRUE' }
VERSION : 0.1
// stored: AutoNumber true, IsIECCheckEnabled false, SetENOAutomatically false, UDAEnableTagReadback false
   VAR_INPUT
      Startup : Bool;
      Root : Bool;
      Scope : String;
   END_VAR
   VAR_IN_OUT
      Access : "FRK_Access";
   END_VAR
   VAR_TEMP
      Index : Int;
      FreeSlot : Int;
   END_VAR
BEGIN

   IF NOT #Startup THEN
       RETURN;
   END_IF;
   #Access.PolicySlot := 0;
   #Access.PolicyLost := FALSE;
   #Access.PolicyLossAlarm := 0;
   #Access.UserLossAlarm := 0;
   IF NOT #Root THEN
       RETURN;
   END_IF;
   #FreeSlot := 0;
   FOR #Index := 1 TO 1 DO
       IF "FRK_AccessPolicies".Rows[#Index].Scope = #Scope THEN
           IF #Access.PolicySlot <> 0 THEN
               #Access.PolicyLost := TRUE;
           ELSE
               #Access.PolicySlot := #Index;
           END_IF;
       ELSIF #FreeSlot = 0 AND NOT "FRK_AccessPolicies".Rows[#Index].Initialized AND "FRK_AccessPolicies".Rows[#Index].Scope = '' AND "FRK_AccessPolicies".Rows[#Index].SchemaVersion = 0 AND "FRK_AccessPolicies".Rows[#Index].Generation = 0 AND "FRK_AccessPolicies".Rows[#Index].Checksum = DWORD#0 THEN
           #FreeSlot := #Index;
       END_IF;
   END_FOR;
   IF #Access.PolicySlot > 0 THEN
       IF NOT #Access.PolicyLost AND "FRK_AccessPolicyValid"(Image := "FRK_AccessPolicies".Rows[#Access.PolicySlot]) THEN
           #Access.Policy := "FRK_AccessPolicies".Rows[#Access.PolicySlot].Policy;
       ELSE
           #Access.PolicyLost := TRUE;
       END_IF;
   ELSIF #FreeSlot > 0 THEN
       #Access.PolicySlot := #FreeSlot;
       "FRK_AccessPolicySave"(Access := #Access,
                              Scope := #Scope);
   ELSE
       #Access.PolicyLost := TRUE;
   END_IF;
   IF #Access.PolicyLost THEN
       // Do not silently reopen actions after losing commissioned policy.
       #Access.Policy := "FRK_AccessStorage".EmptyPolicy;
       FOR #Index := 0 TO 11 DO
           #Access.Policy.Required[#Index] := 4;
       END_FOR;
   END_IF;
END_FUNCTION

FUNCTION "FRK_AccessPolicyCrc" : DWord   // FC55, SCL
{ S7_Optimized_Access := 'TRUE' }
VERSION : 0.1
// stored: AutoNumber true, IsIECCheckEnabled false, SetENOAutomatically false, UDAEnableTagReadback false
   VAR_IN_OUT
      Image : "FRK_AccessPolicyImage";
   END_VAR
   VAR_TEMP
      Work : DWord;
      Index : Int;
      Size : Int;
   END_VAR
BEGIN

   #Work := "FRK_AccessCrcNumber"(Previous := DWORD#16#FFFFFFFF, Value := UINT_TO_UDINT(#Image.SchemaVersion));
   IF #Image.Initialized THEN
       #Work := "FRK_AccessCrcByte"(Previous := #Work, Value := BYTE#1);
   ELSE
       #Work := "FRK_AccessCrcByte"(Previous := #Work, Value := BYTE#0);
   END_IF;
   #Work := "FRK_AccessCrcNumber"(Previous := #Work, Value := #Image.Generation);
   #Size := LEN(#Image.Scope);
   #Work := "FRK_AccessCrcNumber"(Previous := #Work, Value := INT_TO_UDINT(#Size));
   FOR #Index := 1 TO #Size DO
       #Work := "FRK_AccessCrcByte"(Previous := #Work, Value := CHAR_TO_BYTE(#Image.Scope[#Index]));
   END_FOR;
   FOR #Index := 0 TO 11 DO
       #Work := "FRK_AccessCrcNumber"(Previous := #Work, Value := DINT_TO_UDINT(#Image.Policy.Required[#Index]));
   END_FOR;
   #Work := "FRK_AccessCrcNumber"(Previous := #Work, Value := DINT_TO_UDINT(TIME_TO_DINT(#Image.Policy.SessionTimeout)));
   #FRK_AccessPolicyCrc := NOT #Work;
END_FUNCTION

FUNCTION "FRK_AccessPolicySave" : Void   // FC58, SCL
{ S7_Optimized_Access := 'TRUE' }
VERSION : 0.1
// stored: AutoNumber true, IsIECCheckEnabled false, SetENOAutomatically false, UDAEnableTagReadback false
   VAR_INPUT
      Scope : String;
   END_VAR
   VAR_IN_OUT
      Access : "FRK_Access";
   END_VAR
BEGIN

   IF #Access.PolicySlot < 1 OR #Access.PolicySlot > 1 THEN
       RETURN;
   END_IF;
   IF #Scope = '' OR NOT "FRK_AccessPolicyShape"(Policy := #Access.Policy) THEN
       #Access.PolicyLost := TRUE;
       RETURN;
   END_IF;
   "FRK_AccessPolicies".Rows[#Access.PolicySlot].SchemaVersion := 1;
   "FRK_AccessPolicies".Rows[#Access.PolicySlot].Initialized := TRUE;
   "FRK_AccessPolicies".Rows[#Access.PolicySlot].Scope := #Scope;
   "FRK_AccessPolicies".Rows[#Access.PolicySlot].Generation := "FRK_AccessNext"(Previous := "FRK_AccessPolicies".Rows[#Access.PolicySlot].Generation);
   "FRK_AccessPolicies".Rows[#Access.PolicySlot].Policy := #Access.Policy;
   "FRK_AccessPolicies".Rows[#Access.PolicySlot].Checksum := "FRK_AccessPolicyCrc"(Image := "FRK_AccessPolicies".Rows[#Access.PolicySlot]);
END_FUNCTION

FUNCTION "FRK_AccessPolicyShape" : Bool   // FC56, SCL
{ S7_Optimized_Access := 'TRUE' }
VERSION : 0.1
// stored: AutoNumber true, IsIECCheckEnabled false, SetENOAutomatically false, UDAEnableTagReadback false
   VAR_IN_OUT
      Policy : "ST_AccessPolicy";
   END_VAR
   VAR_TEMP
      Index : Int;
   END_VAR
BEGIN

   #FRK_AccessPolicyShape := FALSE;
   IF #Policy.SessionTimeout < T#0ms OR #Policy.SessionTimeout > T#604800000ms THEN
       RETURN;
   END_IF;
   FOR #Index := 0 TO 11 DO
       IF #Policy.Required[#Index] < 0 OR #Policy.Required[#Index] > 4 THEN
           RETURN;
       END_IF;
   END_FOR;
   #FRK_AccessPolicyShape := TRUE;
END_FUNCTION

FUNCTION "FRK_AccessPolicyValid" : Bool   // FC57, SCL
{ S7_Optimized_Access := 'TRUE' }
VERSION : 0.1
// stored: AutoNumber true, IsIECCheckEnabled false, SetENOAutomatically false, UDAEnableTagReadback false
   VAR_IN_OUT
      Image : "FRK_AccessPolicyImage";
   END_VAR
   VAR_TEMP
      Index : Int;
   END_VAR
BEGIN

   #FRK_AccessPolicyValid := FALSE;
   IF NOT #Image.Initialized OR #Image.SchemaVersion <> 1 OR #Image.Scope = '' OR #Image.Generation = 0 OR NOT "FRK_AccessPolicyShape"(Policy := #Image.Policy) THEN
       RETURN;
   END_IF;
   #FRK_AccessPolicyValid := #Image.Checksum = "FRK_AccessPolicyCrc"(Image := #Image);
END_FUNCTION

FUNCTION "FRK_AccessRegisterHash" : Bool   // FC53, SCL
{ S7_Optimized_Access := 'TRUE' }
VERSION : 0.1
// stored: AutoNumber true, IsIECCheckEnabled false, SetENOAutomatically false, UDAEnableTagReadback false
   VAR_INPUT
      Record : "ST_UserRecord";
   END_VAR
   VAR_TEMP
      Slot : Int;
      Index : Int;
   END_VAR
BEGIN

   // Trusted composition/provider seam, never a remote credential editor.
   #FRK_AccessRegisterHash := FALSE;
   IF NOT "FRK_AccessStorage".UsersReady OR #Record.User = '' OR #Record.Level < 0 OR #Record.Level > 4 THEN
       RETURN;
   END_IF;
   #Slot := 0;
   FOR #Index := 1 TO DINT_TO_INT("FRK_LocalUsers".Count) DO
       IF "FRK_LocalUsers".Rows[#Index].User = #Record.User THEN
           #Slot := #Index;
           EXIT;
       END_IF;
   END_FOR;
   IF #Slot = 0 THEN
       IF "FRK_LocalUsers".Count = 16 THEN
           RETURN;
       END_IF;
       "FRK_LocalUsers".Count := "FRK_LocalUsers".Count + 1;
       #Slot := DINT_TO_INT("FRK_LocalUsers".Count);
   END_IF;
   "FRK_LocalUsers".Rows[#Slot] := #Record;
   #FRK_AccessRegisterHash := "FRK_AccessUsersCommit"();
END_FUNCTION

FUNCTION "FRK_AccessStoreBoot" : Void   // FC54, SCL
{ S7_Optimized_Access := 'TRUE' }
VERSION : 0.1
// stored: AutoNumber true, IsIECCheckEnabled false, SetENOAutomatically false, UDAEnableTagReadback false
   VAR_INPUT
      Startup : Bool;
   END_VAR
   VAR_TEMP
      Accepted : Bool;
   END_VAR
BEGIN

   IF NOT #Startup THEN
       RETURN;
   END_IF;
   "FRK_AccessStorage".UsersReady := FALSE;
   "FRK_AccessStorage".UsersLost := FALSE;
   // A virgin image may accept deliberate composition-root provisioning.
   IF NOT "FRK_AccessStorage".UsersCommissioned AND "FRK_LocalUsers".SchemaVersion = 0 AND "FRK_LocalUsers".Generation = 0 AND "FRK_LocalUsers".Checksum = DWORD#0 THEN
       #Accepted := "FRK_AccessUsersCommit"();
       "FRK_AccessStorage".UsersLost := NOT #Accepted;
   ELSIF "FRK_AccessStorage".UsersCommissioned AND "FRK_LocalUsers".SchemaVersion = 1 AND "FRK_LocalUsers".Generation > 0 AND "FRK_AccessUsersShape"() THEN
       "FRK_AccessStorage".UsersReady := "FRK_LocalUsers".Checksum = "FRK_AccessUsersCrc"();
       "FRK_AccessStorage".UsersLost := NOT "FRK_AccessStorage".UsersReady;
   ELSE
       "FRK_AccessStorage".UsersLost := TRUE;
   END_IF;
END_FUNCTION

FUNCTION "FRK_AccessUsersCommit" : Bool   // FC52, SCL
{ S7_Optimized_Access := 'TRUE' }
VERSION : 0.1
// stored: AutoNumber true, IsIECCheckEnabled false, SetENOAutomatically false, UDAEnableTagReadback false
BEGIN

   #FRK_AccessUsersCommit := "FRK_AccessUsersShape"();
   IF NOT #FRK_AccessUsersCommit THEN
       RETURN;
   END_IF;
   "FRK_LocalUsers".SchemaVersion := 1;
   "FRK_LocalUsers".Generation := "FRK_AccessNext"(Previous := "FRK_LocalUsers".Generation);
   "FRK_LocalUsers".Checksum := "FRK_AccessUsersCrc"();
   "FRK_AccessStorage".UsersCommissioned := TRUE;
   "FRK_AccessStorage".UsersReady := TRUE;
   "FRK_AccessStorage".UsersLost := FALSE;
END_FUNCTION

FUNCTION "FRK_AccessUsersCrc" : DWord   // FC50, SCL
{ S7_Optimized_Access := 'TRUE' }
VERSION : 0.1
// stored: AutoNumber true, IsIECCheckEnabled false, SetENOAutomatically false, UDAEnableTagReadback false
   VAR_TEMP
      Work : DWord;
      Slot : Int;
      Index : Int;
      Size : Int;
   END_VAR
BEGIN

   #Work := "FRK_AccessCrcNumber"(Previous := DWORD#16#FFFFFFFF, Value := UINT_TO_UDINT("FRK_LocalUsers".SchemaVersion));
   #Work := "FRK_AccessCrcNumber"(Previous := #Work, Value := "FRK_LocalUsers".Generation);
   #Work := "FRK_AccessCrcNumber"(Previous := #Work, Value := DINT_TO_UDINT("FRK_LocalUsers".Count));
   // Unused rows are included: an altered dormant credential is not ignored.
   FOR #Slot := 1 TO 16 DO
       #Size := LEN("FRK_LocalUsers".Rows[#Slot].User);
       #Work := "FRK_AccessCrcNumber"(Previous := #Work, Value := INT_TO_UDINT(#Size));
       FOR #Index := 1 TO #Size DO
           #Work := "FRK_AccessCrcByte"(Previous := #Work, Value := CHAR_TO_BYTE("FRK_LocalUsers".Rows[#Slot].User[#Index]));
       END_FOR;
       #Work := "FRK_AccessCrcNumber"(Previous := #Work, Value := DINT_TO_UDINT("FRK_LocalUsers".Rows[#Slot].Level));
       FOR #Index := 0 TO 15 DO
           #Work := "FRK_AccessCrcByte"(Previous := #Work, Value := "FRK_LocalUsers".Rows[#Slot].Salt[#Index]);
       END_FOR;
       FOR #Index := 0 TO 31 DO
           #Work := "FRK_AccessCrcByte"(Previous := #Work, Value := "FRK_LocalUsers".Rows[#Slot].PinHash[#Index]);
       END_FOR;
   END_FOR;
   #FRK_AccessUsersCrc := NOT #Work;
END_FUNCTION

FUNCTION "FRK_AccessUsersShape" : Bool   // FC51, SCL
{ S7_Optimized_Access := 'TRUE' }
VERSION : 0.1
// stored: AutoNumber true, IsIECCheckEnabled false, SetENOAutomatically false, UDAEnableTagReadback false
   VAR_TEMP
      Slot : Int;
      Other : Int;
   END_VAR
BEGIN

   #FRK_AccessUsersShape := FALSE;
   IF "FRK_LocalUsers".Count < 0 OR "FRK_LocalUsers".Count > 16 THEN
       RETURN;
   END_IF;
   FOR #Slot := 1 TO DINT_TO_INT("FRK_LocalUsers".Count) DO
       IF "FRK_LocalUsers".Rows[#Slot].User = '' OR "FRK_LocalUsers".Rows[#Slot].Level < 0 OR "FRK_LocalUsers".Rows[#Slot].Level > 4 THEN
           RETURN;
       END_IF;
       FOR #Other := 1 TO #Slot - 1 DO
           IF "FRK_LocalUsers".Rows[#Slot].User = "FRK_LocalUsers".Rows[#Other].User THEN
               RETURN;
           END_IF;
       END_FOR;
   END_FOR;
   #FRK_AccessUsersShape := TRUE;
END_FUNCTION

FUNCTION "FRK_AdoptFault" : Void   // FC9, SCL
{ S7_Optimized_Access := 'TRUE' }
VERSION : 0.1
// stored: AutoNumber true, IsIECCheckEnabled false, SetENOAutomatically false, UDAEnableTagReadback false
   VAR_INPUT
      Diag : "ST_Diagnostic";
   END_VAR
   VAR_IN_OUT
      Core : "FRK_Core";
      Status : "ST_ModuleStatus";
   END_VAR
BEGIN

   IF #Core.Exec = 3 THEN
       RETURN;
   END_IF;
   #Status.Diagnostic := #Diag;
   #Core.Exec := 3;
   #Core.Step := 0;
   #Core.Dispatch := FALSE;
   #Core.DiagTouched := TRUE;
END_FUNCTION

FUNCTION "FRK_AlarmBegin" : Void   // FC30, SCL
{ S7_Optimized_Access := 'TRUE' }
VERSION : 0.1
// stored: AutoNumber true, IsIECCheckEnabled false, SetENOAutomatically false, UDAEnableTagReadback false
   VAR_INPUT
      Startup : Bool;
   END_VAR
   VAR_IN_OUT
      AlarmLog : "FRK_AlarmLog";
   END_VAR
   VAR_TEMP
      Index : Int;
   END_VAR
BEGIN

   FOR #Index := 1 TO 16 DO
       #AlarmLog.Touched[#Index] := FALSE;
       IF #Startup THEN
           #AlarmLog.Active[#Index] := "FRK_UnitScratch".EmptyEvent;
           #AlarmLog.Automatic[#Index] := FALSE;
           #AlarmLog.ComeMs[#Index] := 0;
       END_IF;
   END_FOR;
   IF #Startup THEN
       FOR #Index := 1 TO 64 DO
           #AlarmLog.Ring[#Index] := "FRK_UnitScratch".EmptyEvent;
       END_FOR;
       #AlarmLog.RingHead := 0;
       #AlarmLog.RingUsed := 0;
       #AlarmLog.Truncated := FALSE;
   END_IF;
   "FRK_AlarmRefresh"(AlarmLog := #AlarmLog);
END_FUNCTION

FUNCTION "FRK_AlarmCapture" : Void   // FC36, SCL
{ S7_Optimized_Access := 'TRUE' }
VERSION : 0.1
// stored: AutoNumber true, IsIECCheckEnabled false, SetENOAutomatically false, UDAEnableTagReadback false
   VAR_IN_OUT
      AlarmLog : "FRK_AlarmLog";
      Core : "FRK_Core";
      Status : "ST_ModuleStatus";
   END_VAR
   VAR_TEMP
      Slot : Int;
   END_VAR
BEGIN

   #Slot := #Core.FaultSlot;
   IF #Slot < 1 OR #Slot > 16 THEN
       #Slot := 0;
   ELSIF NOT #AlarmLog.Automatic[#Slot] OR #AlarmLog.Active[#Slot].State <> 1
       OR #AlarmLog.Active[#Slot].SourcePath <> #Status.Diagnostic.SourcePath
       OR #AlarmLog.Active[#Slot].ReasonCode <> #Status.Diagnostic.ReasonCode
       OR #AlarmLog.Active[#Slot].Description <> #Status.Diagnostic.Description THEN
       #Slot := 0;
   END_IF;
   IF #Core.Exec = 3 AND NOT #Core.FaultHandled THEN
       IF #Slot = 0 THEN
           // Adopted first-outs share one active occurrence within this log.
           FOR #Slot := 1 TO 16 DO
               IF #AlarmLog.Automatic[#Slot] AND #AlarmLog.Active[#Slot].State = 1
                   AND #AlarmLog.Active[#Slot].SourcePath = #Status.Diagnostic.SourcePath
                   AND #AlarmLog.Active[#Slot].ReasonCode = #Status.Diagnostic.ReasonCode
                   AND #AlarmLog.Active[#Slot].Description = #Status.Diagnostic.Description THEN
                   EXIT;
               END_IF;
           END_FOR;
           IF #Slot > 16 THEN
               #Slot := "FRK_AlarmRaise"(AlarmLog := #AlarmLog, Diag := #Status.Diagnostic, ResetClass := 1);
           END_IF;
       END_IF;
       IF #Slot > 0 THEN
           #AlarmLog.Automatic[#Slot] := TRUE;
           #AlarmLog.Touched[#Slot] := TRUE;
       END_IF;
       #Core.FaultSlot := #Slot;
   ELSE
       #Core.FaultSlot := 0;
   END_IF;
END_FUNCTION

FUNCTION "FRK_AlarmClose" : Void   // FC32, SCL
{ S7_Optimized_Access := 'TRUE' }
VERSION : 0.1
// stored: AutoNumber true, IsIECCheckEnabled false, SetENOAutomatically false, UDAEnableTagReadback false
   VAR_INPUT
      Slot : Int;
   END_VAR
   VAR_IN_OUT
      AlarmLog : "FRK_AlarmLog";
   END_VAR
BEGIN

   IF #Slot < 1 OR #Slot > 16 THEN
       RETURN;
   END_IF;
   IF #AlarmLog.Active[#Slot].State = 0 THEN
       RETURN;
   END_IF;
   #AlarmLog.Active[#Slot].State := 0;
   IF #AlarmLog.RingHead < 0 OR #AlarmLog.RingHead > 64 THEN
       #AlarmLog.RingHead := 0;
   END_IF;
   #AlarmLog.RingHead := (#AlarmLog.RingHead MOD 64) + 1;
   IF #AlarmLog.RingUsed >= 64 THEN
       #AlarmLog.Truncated := TRUE;
   ELSE
       #AlarmLog.RingUsed := #AlarmLog.RingUsed + 1;
   END_IF;
   #AlarmLog.Ring[#AlarmLog.RingHead] := #AlarmLog.Active[#Slot];
   #AlarmLog.Automatic[#Slot] := FALSE;
   "FRK_AlarmRefresh"(AlarmLog := #AlarmLog);
   "FRK_AlarmNotify"(AlarmLog := #AlarmLog,
                     Ev := #AlarmLog.Ring[#AlarmLog.RingHead]);
END_FUNCTION

FUNCTION "FRK_AlarmEnd" : Void   // FC37, SCL
{ S7_Optimized_Access := 'TRUE' }
VERSION : 0.1
// stored: AutoNumber true, IsIECCheckEnabled false, SetENOAutomatically false, UDAEnableTagReadback false
   VAR_IN_OUT
      AlarmLog : "FRK_AlarmLog";
   END_VAR
   VAR_TEMP
      Slot : Int;
      Gone : Bool;
   END_VAR
BEGIN

   FOR #Slot := 1 TO 16 DO
       IF #AlarmLog.Automatic[#Slot] AND NOT #AlarmLog.Touched[#Slot] THEN
           #Gone := "FRK_AlarmGone"(AlarmLog := #AlarmLog, Slot := #Slot);
       END_IF;
   END_FOR;
END_FUNCTION

FUNCTION "FRK_AlarmGone" : Bool   // FC33, SCL
{ S7_Optimized_Access := 'TRUE' }
VERSION : 0.1
// stored: AutoNumber true, IsIECCheckEnabled false, SetENOAutomatically false, UDAEnableTagReadback false
   VAR_INPUT
      Slot : Int;
   END_VAR
   VAR_IN_OUT
      AlarmLog : "FRK_AlarmLog";
   END_VAR
   VAR_TEMP
      Span : UDInt;
      Stamp : DTL;
      ResultCode : Int;
   END_VAR
BEGIN

   #FRK_AlarmGone := FALSE;
   IF #Slot < 1 OR #Slot > 16 THEN
       RETURN;
   END_IF;
   IF #AlarmLog.Active[#Slot].State <> 1 THEN
       RETURN;
   END_IF;
   #ResultCode := RD_SYS_T(OUT => #Stamp);
   IF #ResultCode = 0 THEN
       #AlarmLog.Active[#Slot].GoneAt := DTL_TO_LDT(#Stamp);
   END_IF;
   #AlarmLog.Active[#Slot].GoneTimeSynchronized := FALSE;
   #Span := "FRK_Elapsed"(NewMs := "FRK_Clock".NowMs, OldMs := #AlarmLog.ComeMs[#Slot]);
   IF #Span > 2147483647 THEN
       #Span := 2147483647;
   END_IF;
   #AlarmLog.Active[#Slot].Duration := DINT_TO_TIME(UDINT_TO_DINT(#Span));
   IF #AlarmLog.Active[#Slot].ResetClass = 0 THEN
       "FRK_AlarmClose"(AlarmLog := #AlarmLog,
                        Slot := #Slot);
   ELSE
       #AlarmLog.Active[#Slot].State := 2;
       #AlarmLog.Automatic[#Slot] := FALSE;
   END_IF;
   #FRK_AlarmGone := TRUE;
END_FUNCTION

FUNCTION "FRK_AlarmMessage" : Void   // FC35, SCL
{ S7_Optimized_Access := 'TRUE' }
VERSION : 0.1
// stored: AutoNumber true, IsIECCheckEnabled false, SetENOAutomatically false, UDAEnableTagReadback false
   VAR_INPUT
      Reason : DInt;
      Description : WString;
      SourcePath : WString;
   END_VAR
   VAR_IN_OUT
      AlarmLog : "FRK_AlarmLog";
   END_VAR
   VAR_TEMP
      Diag : "ST_Diagnostic";
      Slot : Int;
      Gone : Bool;
   END_VAR
BEGIN

   #Diag := "FRK_UnitScratch".EmptyDiagnostic;
   #Diag.ReasonCode := #Reason;
   #Diag.Description := #Description;
   #Diag.SourcePath := #SourcePath;
   #Diag.Severity := 0;
   #Diag.Category := 2;
   #Slot := "FRK_AlarmRaise"(AlarmLog := #AlarmLog, Diag := #Diag, ResetClass := 0);
   IF #Slot > 0 THEN
       #Gone := "FRK_AlarmGone"(AlarmLog := #AlarmLog, Slot := #Slot);
   END_IF;
END_FUNCTION

FUNCTION "FRK_AlarmNotify" : Void   // FC28, SCL
{ S7_Optimized_Access := 'TRUE' }
VERSION : 0.1
// Core 8.3: one owning active list / closed ring, with optional event callback.
// stored: AutoNumber true, IsIECCheckEnabled false, SetENOAutomatically false, UDAEnableTagReadback false
   VAR_INPUT
      Ev : "ST_AlarmEvent";
   END_VAR
   VAR_IN_OUT
      AlarmLog : "FRK_AlarmLog";
   END_VAR
BEGIN

   RETURN; // No event sink supplied by the composition declaration.
END_FUNCTION

FUNCTION "FRK_AlarmOperatorReset" : Void   // FC34, SCL
{ S7_Optimized_Access := 'TRUE' }
VERSION : 0.1
// stored: AutoNumber true, IsIECCheckEnabled false, SetENOAutomatically false, UDAEnableTagReadback false
   VAR_IN_OUT
      AlarmLog : "FRK_AlarmLog";
   END_VAR
   VAR_TEMP
      Slot : Int;
      Gone : Bool;
      Stamp : DTL;
      ResultCode : Int;
   END_VAR
BEGIN

   FOR #Slot := 1 TO 16 DO
       IF #AlarmLog.Active[#Slot].State <> 0 AND #AlarmLog.Active[#Slot].ResetClass = 1 THEN
           IF #AlarmLog.Active[#Slot].State = 1 THEN
               #Gone := "FRK_AlarmGone"(AlarmLog := #AlarmLog, Slot := #Slot);
           END_IF;
           #ResultCode := RD_SYS_T(OUT => #Stamp);
           IF #ResultCode = 0 THEN
               #AlarmLog.Active[#Slot].ResetAt := DTL_TO_LDT(#Stamp);
           END_IF;
           #AlarmLog.Active[#Slot].ResetTimeSynchronized := FALSE;
           "FRK_AlarmClose"(AlarmLog := #AlarmLog,
                            Slot := #Slot);
       END_IF;
   END_FOR;
END_FUNCTION

FUNCTION "FRK_AlarmRaise" : Int   // FC31, SCL
{ S7_Optimized_Access := 'TRUE' }
VERSION : 0.1
// stored: AutoNumber true, IsIECCheckEnabled false, SetENOAutomatically false, UDAEnableTagReadback false
   VAR_INPUT
      Diag : "ST_Diagnostic";
      ResetClass : DInt;
   END_VAR
   VAR_IN_OUT
      AlarmLog : "FRK_AlarmLog";
   END_VAR
   VAR_TEMP
      Slot : Int;
      Stamp : DTL;
      ResultCode : Int;
      Rational : "ST_Diagnostic";
   END_VAR
BEGIN

   #FRK_AlarmRaise := 0;
   IF #ResetClass < 0 OR #ResetClass > 1
       OR #Diag.Severity < 0 OR #Diag.Severity > 2
       OR #Diag.Category < 0 OR #Diag.Category > 2
       OR #Diag.SourcePath = WSTRING#'' OR #Diag.Description = WSTRING#'' THEN
       RETURN;
   END_IF;
   FOR #Slot := 1 TO 16 DO
       IF #AlarmLog.Active[#Slot].State = 0 THEN
           #Rational := #Diag;
           "FRK_Rationalize"(Diag := #Rational);
           #AlarmLog.Active[#Slot] := "FRK_UnitScratch".EmptyEvent;
           #AlarmLog.Active[#Slot].ReasonCode := #Rational.ReasonCode;
           #AlarmLog.Active[#Slot].Description := #Rational.Description;
           #AlarmLog.Active[#Slot].SourcePath := #Rational.SourcePath;
           #AlarmLog.Active[#Slot].IoTag := #Rational.IoTag;
           #AlarmLog.Active[#Slot].IoAddress := #Rational.IoAddress;
           #AlarmLog.Active[#Slot].Severity := #Rational.Severity;
           #AlarmLog.Active[#Slot].Category := #Rational.Category;
           #AlarmLog.Active[#Slot].ResetClass := #ResetClass;
           #AlarmLog.Active[#Slot].State := 1;
           #AlarmLog.ComeMs[#Slot] := "FRK_Clock".NowMs;
           #AlarmLog.Automatic[#Slot] := FALSE;
           #AlarmLog.Touched[#Slot] := FALSE;
           #ResultCode := RD_SYS_T(OUT => #Stamp);
           IF #ResultCode = 0 THEN
               #AlarmLog.Active[#Slot].ComeAt := DTL_TO_LDT(#Stamp);
           END_IF;
           // The UTC source has no proven synchronization witness yet.
           #AlarmLog.Active[#Slot].ComeTimeSynchronized := FALSE;
           "FRK_AlarmRefresh"(AlarmLog := #AlarmLog);
           "FRK_AlarmNotify"(AlarmLog := #AlarmLog,
                             Ev := #AlarmLog.Active[#Slot]);
           #FRK_AlarmRaise := #Slot;
           RETURN;
       END_IF;
   END_FOR;
   #AlarmLog.Truncated := TRUE;
END_FUNCTION

FUNCTION "FRK_AlarmRefresh" : Void   // FC29, SCL
{ S7_Optimized_Access := 'TRUE' }
VERSION : 0.1
// stored: AutoNumber true, IsIECCheckEnabled false, SetENOAutomatically false, UDAEnableTagReadback false
   VAR_IN_OUT
      AlarmLog : "FRK_AlarmLog";
   END_VAR
   VAR_TEMP
      Index : Int;
   END_VAR
BEGIN

   #AlarmLog.NActive := 0;
   #AlarmLog.Blocking := FALSE;
   FOR #Index := 1 TO 16 DO
       IF #AlarmLog.Active[#Index].State <> 0 THEN
           #AlarmLog.NActive := #AlarmLog.NActive + 1;
           IF #AlarmLog.Active[#Index].ResetClass = 1 THEN
               #AlarmLog.Blocking := TRUE;
           END_IF;
       END_IF;
   END_FOR;
END_FUNCTION

FUNCTION "FRK_AlarmTreeBlocking" : Bool   // FC38, SCL
{ S7_Optimized_Access := 'TRUE' }
VERSION : 0.1
// stored: AutoNumber true, IsIECCheckEnabled false, SetENOAutomatically false, UDAEnableTagReadback false
   VAR_INPUT
      Owner : DInt;
   END_VAR
   VAR_TEMP
      Index : DInt;
      Ancestor : DInt;
      Depth : DInt;
   END_VAR
BEGIN

   #FRK_AlarmTreeBlocking := TRUE;
   IF "FRK_Registry".Fault OR #Owner < 1 OR #Owner > "FRK_Registry".Count OR "FRK_Registry".Count > 4 THEN
       RETURN;
   END_IF;
   FOR #Index := 1 TO "FRK_Registry".Count DO
       IF "FRK_Registry".Rows[#Index].AlarmBlocking THEN
           #Ancestor := #Index;
           FOR #Depth := 1 TO 4 DO
               IF #Ancestor = #Owner THEN
                   RETURN;
               END_IF;
               IF #Ancestor = 0 THEN
                   EXIT;
               END_IF;
               IF #Ancestor < 1 OR #Ancestor > "FRK_Registry".Count THEN
                   RETURN;
               END_IF;
               #Ancestor := "FRK_Registry".Rows[#Ancestor].Parent;
           END_FOR;
           IF #Depth > 4 AND #Ancestor <> 0 THEN
               RETURN;
           END_IF;
       END_IF;
   END_FOR;
   #FRK_AlarmTreeBlocking := FALSE;
END_FUNCTION

FUNCTION "FRK_Begin" : Void   // FC15, SCL
{ S7_Optimized_Access := 'TRUE' }
VERSION : 0.1
// stored: AutoNumber true, IsIECCheckEnabled false, SetENOAutomatically false, UDAEnableTagReadback false
   VAR_INPUT
      Execute : Bool;
      Abort : Bool;
      Command : DInt;
   END_VAR
   VAR_IN_OUT
      Core : "FRK_Core";
      Status : "ST_ModuleStatus";
   END_VAR
BEGIN

   #Core.EvInit := NOT #Core.Initialized;
   #Core.Initialized := TRUE;
   #Core.EvCommandStart := FALSE;
   #Core.EvAbort := FALSE;
   #Core.EvAbortInError := FALSE;
   #Core.HoldReq := FALSE;
   #Core.DiagTouched := FALSE;
   #Core.FaultHandled := FALSE;
   #Core.HookResult := 0;
   IF NOT #Execute AND (#Core.Armed OR #Core.ReleasePending) AND (#Core.Exec = 2 OR #Core.Exec = 3 OR #Core.Exec = 4) THEN
       #Core.Exec := 0;
       #Core.Armed := FALSE;
       #Core.HoldReason := 0;
       "FRK_ClearDiag"(Status := #Status);
   END_IF;
   IF #Execute AND NOT #Core.ExecPrev AND (#Core.Exec = 0 OR (#Core.Exec = 3 AND NOT #Core.Armed)) THEN
       #Core.Exec := 1;
       #Core.Armed := TRUE;
       #Core.Command := #Command;
       #Core.Step := 10;
       #Core.StartMs := "FRK_Clock".NowMs;
       #Core.LastNowMs := "FRK_Clock".NowMs;
       #Core.ActiveMs := 0;
       #Core.TimeoutMs := 0;
       #Core.CommandLabel := '';
       #Core.TimingOpen := TRUE;
       #Core.Held := FALSE;
       #Core.HoldReason := 0;
       "FRK_ClearDiag"(Status := #Status);
       #Core.EvCommandStart := TRUE;
   END_IF;
   #Core.DeltaMs := "FRK_Elapsed"(NewMs := "FRK_Clock".NowMs, OldMs := #Core.LastNowMs);
   #Core.LastNowMs := "FRK_Clock".NowMs;
   #Core.ExecPrev := #Execute;
   #Core.Dispatch := #Core.Exec = 1;
END_FUNCTION

FUNCTION "FRK_Capture_CylinderCM" : Void   // FC152, SCL
{ S7_Optimized_Access := 'TRUE' }
VERSION : 0.1
// stored: AutoNumber true, IsIECCheckEnabled false, SetENOAutomatically false, UDAEnableTagReadback false
   VAR_IN_OUT
      Module : "FB_CylinderCM";
      AlarmLog : "FRK_AlarmLog";
   END_VAR
BEGIN

   "FRK_AlarmCapture"(AlarmLog := #AlarmLog,
                      Core := #Module.Core,
                      Status := #Module.Status);
END_FUNCTION

FUNCTION "FRK_CfgDef_CylinderCM" : Void   // FC147, SCL
{ S7_Optimized_Access := 'TRUE' }
VERSION : 0.1
// stored: AutoNumber true, IsIECCheckEnabled false, SetENOAutomatically false, UDAEnableTagReadback false
   VAR_INPUT
      FieldIndex : Int;
   END_VAR
BEGIN

   "FRK_ConfigScratch".Entry := "FRK_ConfigScratch".Blank;
END_FUNCTION

FUNCTION "FRK_CfgDef_PressDemoUnit" : Void   // FC173, SCL
{ S7_Optimized_Access := 'TRUE' }
VERSION : 0.1
// stored: AutoNumber true, IsIECCheckEnabled false, SetENOAutomatically false, UDAEnableTagReadback false
   VAR_INPUT
      FieldIndex : Int;
   END_VAR
BEGIN

